  MoveL 2059 to (-200, -12.5, 57) mm, rotated rx 180 ry 0 rz 180 deg; joints [-15.333, -59.757, 128.123, 163.566, 69.173, -84.013]
  MoveL 2060 to (0, -12.5, 57) mm, rotated rx 180 ry 0 rz 180 deg; joints [-13.182, -51.64, 111.998, 164.918, 61.214, -82.606]
  MoveL 2061 to (0, -11.9, 57) mm, rotated rx 180 ry 0 rz 180 deg; joints [-13.182, -51.608, 111.999, 164.923, 61.246, -82.616]
  MoveL 2062 to (-200, -11.9, 57) mm, rotated rx 180 ry 0 rz 180 deg; joints [-15.333, -59.718, 128.125, 163.57, 69.212, -84.025]
  MoveL 2063 to (-200, -11.3, 57) mm, rotated rx 180 ry 0 rz 180 deg; joints [-15.333, -59.679, 128.126, 163.574, 69.251, -84.038]
  MoveL 2064 to (0, -11.3, 57) mm, rotated rx 180 ry 0 rz 180 deg; joints [-13.182, -51.576, 112.001, 164.927, 61.278, -82.626]
  MoveL 2065 to (0, -10.7, 57) mm, rotated rx 180 ry 0 rz 180 deg; joints [-13.182, -51.544, 112.002, 164.932, 61.31, -82.636]
  MoveL 2066 to (-200, -10.7, 57) mm, rotated rx 180 ry 0 rz 180 deg; joints [-15.333, -59.64, 128.127, 163.579, 69.289, -84.05]
  MoveL 2067 to (-200, -10.1, 57) mm, rotated rx 180 ry 0 rz 180 deg; joints [-15.333, -59.601, 128.129, 163.583, 69.328, -84.062]
  MoveL 2068 to (0, -10.1, 57) mm, rotated rx 180 ry 0 rz 180 deg; joints [-13.182, -51.512, 112.003, 164.937, 61.341, -82.645]
  MoveL 2069 to (0, -9.5, 57) mm, rotated rx 180 ry 0 rz 180 deg; joints [-13.182, -51.48, 112.004, 164.942, 61.373, -82.655]
  MoveL 2070 to (-200, -9.5, 57) mm, rotated rx 180 ry 0 rz 180 deg; joints [-15.333, -59.561, 128.13, 163.587, 69.367, -84.074]
  MoveL 2071 to (-200, -8.9, 57) mm, rotated rx 180 ry 0 rz 180 deg; joints [-15.333, -59.522, 128.131, 163.592, 69.406, -84.086]
  MoveL 2072 to (0, -8.9, 57) mm, rotated rx 180 ry 0 rz 180 deg; joints [-13.182, -51.449, 112.005, 164.946, 61.405, -82.665]
  MoveL 2073 to (0, -8.3, 57) mm, rotated rx 180 ry 0 rz 180 deg; joints [-13.182, -51.417, 112.006, 164.951, 61.437, -82.675]
  MoveL 2074 to (-200, -8.3, 57) mm, rotated rx 180 ry 0 rz 180 deg; joints [-15.333, -59.483, 128.132, 163.596, 69.444, -84.098]
  MoveL 2075 to (-200, -7.7, 57) mm, rotated rx 180 ry 0 rz 180 deg; joints [-15.333, -59.444, 128.133, 163.6, 69.483, -84.111]
  MoveL 2076 to (0, -7.7, 57) mm, rotated rx 180 ry 0 rz 180 deg; joints [-13.182, -51.385, 112.007, 164.956, 61.469, -82.684]
  MoveL 2077 to (0, -7.1, 57) mm, rotated rx 180 ry 0 rz 180 deg; joints [-13.182, -51.353, 112.008, 164.96, 61.501, -82.694]
  MoveL 2078 to (-200, -7.1, 57) mm, rotated rx 180 ry 0 rz 180 deg; joints [-15.333, -59.405, 128.135, 163.604, 69.522, -84.123]
  MoveL 2079 to (-200, -6.5, 57) mm, rotated rx 180 ry 0 rz 180 deg; joints [-15.333, -59.366, 128.136, 163.609, 69.56, -84.135]
  MoveL 2080 to (0, -6.5, 57) mm, rotated rx 180 ry 0 rz 180 deg; joints [-13.182, -51.321, 112.009, 164.965, 61.533, -82.704]
  MoveL 2081 to (0, -5.9, 57) mm, rotated rx 180 ry 0 rz 180 deg; joints [-13.182, -51.289, 112.01, 164.969, 61.564, -82.714]
  MoveL 2082 to (-200, -5.9, 57) mm, rotated rx 180 ry 0 rz 180 deg; joints [-15.333, -59.327, 128.137, 163.613, 69.599, -84.147]
  MoveL 2083 to (-200, -5.3, 57) mm, rotated rx 180 ry 0 rz 180 deg; joints [-15.333, -59.287, 128.138, 163.617, 69.637, -84.159]
  MoveL 2084 to (0, -5.3, 57) mm, rotated rx 180 ry 0 rz 180 deg; joints [-13.182, -51.257, 112.011, 164.974, 61.596, -82.723]
  MoveL 2085 to (0, -4.7, 57) mm, rotated rx 180 ry 0 rz 180 deg; joints [-13.182, -51.225, 112.012, 164.979, 61.628, -82.733]
  MoveL 2086 to (-200, -4.7, 57) mm, rotated rx 180 ry 0 rz 180 deg; joints [-15.333, -59.248, 128.139, 163.621, 69.676, -84.171]
  MoveL 2087 to (-200, -4.1, 57) mm, rotated rx 180 ry 0 rz 180 deg; joints [-15.333, -59.209, 128.14, 163.626, 69.715, -84.183]
  MoveL 2088 to (0, -4.1, 57) mm, rotated rx 180 ry 0 rz 180 deg; joints [-13.182, -51.193, 112.013, 164.983, 61.66, -82.743]
  MoveL 2089 to (0, -3.5, 57) mm, rotated rx 180 ry 0 rz 180 deg; joints [-13.182, -51.161, 112.014, 164.988, 61.692, -82.752]
  MoveL 2090 to (-200, -3.5, 57) mm, rotated rx 180 ry 0 rz 180 deg; joints [-15.333, -59.17, 128.141, 163.63, 69.753, -84.195]
  MoveL 2091 to (-200, -2.9, 57) mm, rotated rx 180 ry 0 rz 180 deg; joints [-15.333, -59.13, 128.142, 163.634, 69.792, -84.207]
  MoveL 2092 to (0, -2.9, 57) mm, rotated rx 180 ry 0 rz 180 deg; joints [-13.182, -51.129, 112.015, 164.992, 61.723, -82.762]
  MoveL 2093 to (0, -2.3, 57) mm, rotated rx 180 ry 0 rz 180 deg; joints [-13.182, -51.097, 112.015, 164.997, 61.755, -82.772]
  MoveL 2094 to (-200, -2.3, 57) mm, rotated rx 180 ry 0 rz 180 deg; joints [-15.333, -59.091, 128.142, 163.638, 69.83, -84.22]
  MoveL 2095 to (-200, -1.7, 57) mm, rotated rx 180 ry 0 rz 180 deg; joints [-15.333, -59.052, 128.143, 163.642, 69.869, -84.232]
  MoveL 2096 to (0, -1.7, 57) mm, rotated rx 180 ry 0 rz 180 deg; joints [-13.182, -51.064, 112.016, 165.002, 61.787, -82.781]
  MoveL 2097 to (0, -1.1, 57) mm, rotated rx 180 ry 0 rz 180 deg; joints [-13.182, -51.032, 112.017, 165.006, 61.818, -82.791]
  MoveL 2098 to (-200, -1.1, 57) mm, rotated rx 180 ry 0 rz 180 deg; joints [-15.333, -59.012, 128.144, 163.646, 69.907, -84.244]
  MoveL 2099 to (-200, -0.5, 57) mm, rotated rx 180 ry 0 rz 180 deg; joints [-15.333, -58.973, 128.145, 163.651, 69.946, -84.256]
  MoveL 2100 to (0, -0.5, 57) mm, rotated rx 180 ry 0 rz 180 deg; joints [-13.182, -51, 112.017, 165.011, 61.85, -82.801]
  MoveL 2101 to (0, 0, 57) mm, rotated rx 180 ry 0 rz 180 deg; joints [-13.182, -50.974, 112.018, 165.014, 61.876, -82.809]
  MoveL 2102 to (-200, 0, 57) mm, rotated rx 180 ry 0 rz 180 deg; joints [-15.333, -58.94, 128.145, 163.654, 69.978, -84.266]
  MoveL 2103 to (-200, 0, 57.4) mm, rotated rx 180 ry 0 rz 180 deg; joints [-15.351, -58.936, 128.137, 163.634, 69.976, -84.258]
  MoveL 2104 to (0, 0, 57.4) mm, rotated rx 180 ry 0 rz 180 deg; joints [-13.198, -50.97, 112.01, 164.996, 61.875, -82.799]
  MoveL 2105 to (0, -0.6, 57.4) mm, rotated rx 180 ry 0 rz 180 deg; joints [-13.198, -51.002, 112.009, 164.992, 61.843, -82.789]
  MoveL 2106 to (-200, -0.6, 57.4) mm, rotated rx 180 ry 0 rz 180 deg; joints [-15.351, -58.975, 128.136, 163.63, 69.937, -84.246]
  MoveL 2107 to (-200, -1.2, 57.4) mm, rotated rx 180 ry 0 rz 180 deg; joints [-15.351, -59.015, 128.135, 163.626, 69.899, -84.234]
  MoveL 2108 to (0, -1.2, 57.4) mm, rotated rx 180 ry 0 rz 180 deg; joints [-13.198, -51.034, 112.009, 164.987, 61.811, -82.78]
  MoveL 2109 to (0, -1.8, 57.4) mm, rotated rx 180 ry 0 rz 180 deg; joints [-13.198, -51.066, 112.008, 164.982, 61.78, -82.77]
  MoveL 2110 to (-200, -1.8, 57.4) mm, rotated rx 180 ry 0 rz 180 deg; joints [-15.351, -59.054, 128.135, 163.622, 69.86, -84.222]
  MoveL 2111 to (-200, -2.4, 57.4) mm, rotated rx 180 ry 0 rz 180 deg; joints [-15.351, -59.093, 128.134, 163.618, 69.822, -84.21]
  MoveL 2112 to (0, -2.4, 57.4) mm, rotated rx 180 ry 0 rz 180 deg; joints [-13.198, -51.098, 112.007, 164.978, 61.748, -82.76]
  MoveL 2113 to (0, -3, 57.4) mm, rotated rx 180 ry 0 rz 180 deg; joints [-13.198, -51.13, 112.006, 164.973, 61.716, -82.751]
  MoveL 2114 to (-200, -3, 57.4) mm, rotated rx 180 ry 0 rz 180 deg; joints [-15.351, -59.133, 128.133, 163.614, 69.783, -84.198]
  MoveL 2115 to (-200, -3.6, 57.4) mm, rotated rx 180 ry 0 rz 180 deg; joints [-15.351, -59.172, 128.132, 163.609, 69.744, -84.185]
  MoveL 2116 to (0, -3.6, 57.4) mm, rotated rx 180 ry 0 rz 180 deg; joints [-13.198, -51.162, 112.006, 164.969, 61.684, -82.741]
  MoveL 2117 to (0, -4.2, 57.4) mm, rotated rx 180 ry 0 rz 180 deg; joints [-13.198, -51.194, 112.005, 164.964, 61.653, -82.731]
  MoveL 2118 to (-200, -4.2, 57.4) mm, rotated rx 180 ry 0 rz 180 deg; joints [-15.351, -59.211, 128.131, 163.605, 69.706, -84.173]
  MoveL 2119 to (-200, -4.8, 57.4) mm, rotated rx 180 ry 0 rz 180 deg; joints [-15.351, -59.25, 128.13, 163.601, 69.667, -84.161]
  MoveL 2120 to (0, -4.8, 57.4) mm, rotated rx 180 ry 0 rz 180 deg; joints [-13.198, -51.226, 112.004, 164.96, 61.621, -82.722]
  MoveL 2121 to (0, -5.4, 57.4) mm, rotated rx 180 ry 0 rz 180 deg; joints [-13.198, -51.258, 112.003, 164.955, 61.589, -82.712]
  MoveL 2122 to (-200, -5.4, 57.4) mm, rotated rx 180 ry 0 rz 180 deg; joints [-15.351, -59.29, 128.129, 163.597, 69.629, -84.149]
  MoveL 2123 to (-200, -6, 57.4) mm, rotated rx 180 ry 0 rz 180 deg; joints [-15.351, -59.329, 128.128, 163.593, 69.59, -84.137]
  MoveL 2124 to (0, -6, 57.4) mm, rotated rx 180 ry 0 rz 180 deg; joints [-13.198, -51.29, 112.002, 164.95, 61.557, -82.702]
  MoveL 2125 to (0, -6.6, 57.4) mm, rotated rx 180 ry 0 rz 180 deg; joints [-13.198, -51.322, 112.001, 164.946, 61.525, -82.693]
  MoveL 2126 to (-200, -6.6, 57.4) mm, rotated rx 180 ry 0 rz 180 deg; joints [-15.351, -59.368, 128.127, 163.588, 69.551, -84.125]
  MoveL 2127 to (-200, -7.2, 57.4) mm, rotated rx 180 ry 0 rz 180 deg; joints [-15.351, -59.407, 128.126, 163.584, 69.513, -84.113]
  MoveL 2128 to (0, -7.2, 57.4) mm, rotated rx 180 ry 0 rz 180 deg; joints [-13.198, -51.354, 112, 164.941, 61.494, -82.683]
  MoveL 2129 to (0, -7.8, 57.4) mm, rotated rx 180 ry 0 rz 180 deg; joints [-13.198, -51.386, 111.999, 164.936, 61.462, -82.673]
  MoveL 2130 to (-200, -7.8, 57.4) mm, rotated rx 180 ry 0 rz 180 deg; joints [-15.351, -59.446, 128.125, 163.58, 69.474, -84.101]
  MoveL 2131 to (-200, -8.4, 57.4) mm, rotated rx 180 ry 0 rz 180 deg; joints [-15.351, -59.486, 128.124, 163.575, 69.436, -84.088]
  MoveL 2132 to (0, -8.4, 57.4) mm, rotated rx 180 ry 0 rz 180 deg; joints [-13.198, -51.418, 111.998, 164.932, 61.43, -82.663]
  MoveL 2133 to (0, -9, 57.4) mm, rotated rx 180 ry 0 rz 180 deg; joints [-13.198, -51.45, 111.997, 164.927, 61.398, -82.654]
  MoveL 2134 to (-200, -9, 57.4) mm, rotated rx 180 ry 0 rz 180 deg; joints [-15.351, -59.525, 128.123, 163.571, 69.397, -84.076]
  MoveL 2135 to (-200, -9.6, 57.4) mm, rotated rx 180 ry 0 rz 180 deg; joints [-15.351, -59.564, 128.121, 163.567, 69.358, -84.064]
  MoveL 2136 to (0, -9.6, 57.4) mm, rotated rx 180 ry 0 rz 180 deg; joints [-13.198, -51.482, 111.996, 164.922, 61.366, -82.644]
  MoveL 2137 to (0, -10.2, 57.4) mm, rotated rx 180 ry 0 rz 180 deg; joints [-13.198, -51.514, 111.995, 164.918, 61.334, -82.634]
  MoveL 2138 to (-200, -10.2, 57.4) mm, rotated rx 180 ry 0 rz 180 deg; joints [-15.351, -59.603, 128.12, 163.563, 69.319, -84.052]
  MoveL 2139 to (-200, -10.8, 57.4) mm, rotated rx 180 ry 0 rz 180 deg; joints [-15.351, -59.642, 128.119, 163.558, 69.281, -84.04]
  MoveL 2140 to (0, -10.8, 57.4) mm, rotated rx 180 ry 0 rz 180 deg; joints [-13.198, -51.546, 111.994, 164.913, 61.302, -82.624]
  MoveL 2141 to (0, -11.4, 57.4) mm, rotated rx 180 ry 0 rz 180 deg; joints [-13.198, -51.577, 111.992, 164.908, 61.27, -82.614]
  MoveL 2142 to (-200, -11.4, 57.4) mm, rotated rx 180 ry 0 rz 180 deg; joints [-15.351, -59.681, 128.117, 163.554, 69.242, -84.027]
  MoveL 2143 to (-200, -12, 57.4) mm, rotated rx 180 ry 0 rz 180 deg; joints [-15.351, -59.72, 128.116, 163.55, 69.203, -84.015]
  MoveL 2144 to (0, -12, 57.4) mm, rotated rx 180 ry 0 rz 180 deg; joints [-13.198, -51.609, 111.991, 164.903, 61.239, -82.605]
  MoveL 2145 to (0, -12.6, 57.4) mm, rotated rx 180 ry 0 rz 180 deg; joints [-13.198, -51.641, 111.99, 164.899, 61.207, -82.595]
  MoveL 2146 to (-200, -12.6, 57.4) mm, rotated rx 180 ry 0 rz 180 deg; joints [-15.351, -59.759, 128.115, 163.545, 69.164, -84.003]
  MoveL 2147 to (-200, -13.2, 57.4) mm, rotated rx 180 ry 0 rz 180 deg; joints [-15.351, -59.798, 128.113, 163.541, 69.126, -83.991]
  MoveL 2148 to (0, -13.2, 57.4) mm, rotated rx 180 ry 0 rz 180 deg; joints [-13.198, -51.673, 111.989, 164.894, 61.175, -82.585]
  MoveL 2149 to (0, -13.8, 57.4) mm, rotated rx 180 ry 0 rz 180 deg; joints [-13.198, -51.705, 111.987, 164.889, 61.143, -82.575]
  MoveL 2150 to (-200, -13.8, 57.4) mm, rotated rx 180 ry 0 rz 180 deg; joints [-15.351, -59.837, 128.112, 163.537, 69.087, -83.978]
  MoveL 2151 to (-200, -14.4, 57.4) mm, rotated rx 180 ry 0 rz 180 deg; joints [-15.351, -59.876, 128.11, 163.532, 69.048, -83.966]
  MoveL 2152 to (0, -14.4, 57.4) mm, rotated rx 180 ry 0 rz 180 deg; joints [-13.198, -51.736, 111.986, 164.884, 61.111, -82.565]
  MoveL 2153 to (0, -15, 57.4) mm, rotated rx 180 ry 0 rz 180 deg; joints [-13.198, -51.768, 111.985, 164.88, 61.079, -82.555]
  MoveL 2154 to (-200, -15, 57.4) mm, rotated rx 180 ry 0 rz 180 deg; joints [-15.351, -59.915, 128.109, 163.528, 69.009, -83.954]
  MoveL 2155 to (-200, -15.6, 57.4) mm, rotated rx 180 ry 0 rz 180 deg; joints [-15.351, -59.954, 128.107, 163.523, 68.97, -83.941]
  MoveL 2156 to (0, -15.6, 57.4) mm, rotated rx 180 ry 0 rz 180 deg; joints [-13.198, -51.8, 111.983, 164.875, 61.047, -82.545]
  MoveL 2157 to (0, -16.2, 57.4) mm, rotated rx 180 ry 0 rz 180 deg; joints [-13.198, -51.832, 111.982, 164.87, 61.015, -82.535]
  MoveL 2158 to (-200, -16.2, 57.4) mm, rotated rx 180 ry 0 rz 180 deg; joints [-15.351, -59.993, 128.106, 163.519, 68.932, -83.929]
  MoveL 2159 to (-200, -16.8, 57.4) mm, rotated rx 180 ry 0 rz 180 deg; joints [-15.351, -60.032, 128.104, 163.514, 68.893, -83.917]
  MoveL 2160 to (0, -16.8, 57.4) mm, rotated rx 180 ry 0 rz 180 deg; joints [-13.198, -51.863, 111.98, 164.865, 60.983, -82.526]
  MoveL 2161 to (0, -17.4, 57.4) mm, rotated rx 180 ry 0 rz 180 deg; joints [-13.198, -51.895, 111.979, 164.861, 60.951, -82.516]
  MoveL 2162 to (-200, -17.4, 57.4) mm, rotated rx 180 ry 0 rz 180 deg; joints [-15.351, -60.071, 128.102, 163.51, 68.854, -83.905]
  MoveL 2163 to (-200, -18, 57.4) mm, rotated rx 180 ry 0 rz 180 deg; joints [-15.351, -60.11, 128.101, 163.506, 68.815, -83.892]
  MoveL 2164 to (0, -18, 57.4) mm, rotated rx 180 ry 0 rz 180 deg; joints [-13.198, -51.927, 111.977, 164.856, 60.919, -82.506]
  MoveL 2165 to (0, -18.6, 57.4) mm, rotated rx 180 ry 0 rz 180 deg; joints [-13.198, -51.959, 111.976, 164.851, 60.886, -82.496]
  MoveL 2166 to (-200, -18.6, 57.4) mm, rotated rx 180 ry 0 rz 180 deg; joints [-15.351, -60.148, 128.099, 163.501, 68.776, -83.88]
  MoveL 2167 to (-200, -19.2, 57.4) mm, rotated rx 180 ry 0 rz 180 deg; joints [-15.351, -60.187, 128.097, 163.497, 68.737, -83.867]
  MoveL 2168 to (0, -19.2, 57.4) mm, rotated rx 180 ry 0 rz 180 deg; joints [-13.198, -51.99, 111.974, 164.846, 60.854, -82.486]
  MoveL 2169 to (0, -19.8, 57.4) mm, rotated rx 180 ry 0 rz 180 deg; joints [-13.198, -52.022, 111.972, 164.841, 60.822, -82.476]
  MoveL 2170 to (-200, -19.8, 57.4) mm, rotated rx 180 ry 0 rz 180 deg; joints [-15.351, -60.226, 128.095, 163.492, 68.698, -83.855]
  MoveL 2171 to (-200, -20.4, 57.4) mm, rotated rx 180 ry 0 rz 180 deg; joints [-15.351, -60.265, 128.094, 163.488, 68.659, -83.843]
  MoveL 2172 to (0, -20.4, 57.4) mm, rotated rx 180 ry 0 rz 180 deg; joints [-13.198, -52.053, 111.971, 164.836, 60.79, -82.466]
  MoveL 2173 to (0, -21, 57.4) mm, rotated rx 180 ry 0 rz 180 deg; joints [-13.198, -52.085, 111.969, 164.831, 60.758, -82.456]
  MoveL 2174 to (-200, -21, 57.4) mm, rotated rx 180 ry 0 rz 180 deg; joints [-15.351, -60.304, 128.092, 163.483, 68.62, -83.83]
  MoveL 2175 to (-200, -21.6, 57.4) mm, rotated rx 180 ry 0 rz 180 deg; joints [-15.351, -60.342, 128.09, 163.479, 68.581, -83.818]
  MoveL 2176 to (0, -21.6, 57.4) mm, rotated rx 180 ry 0 rz 180 deg; joints [-13.198, -52.117, 111.967, 164.827, 60.726, -82.446]
  MoveL 2177 to (0, -22.2, 57.4) mm, rotated rx 180 ry 0 rz 180 deg; joints [-13.198, -52.148, 111.966, 164.822, 60.694, -82.436]
  MoveL 2178 to (-200, -22.2, 57.4) mm, rotated rx 180 ry 0 rz 180 deg; joints [-15.351, -60.381, 128.088, 163.474, 68.542, -83.805]
  MoveL 2179 to (-200, -22.8, 57.4) mm, rotated rx 180 ry 0 rz 180 deg; joints [-15.351, -60.42, 128.086, 163.469, 68.503, -83.793]
  MoveL 2180 to (0, -22.8, 57.4) mm, rotated rx 180 ry 0 rz 180 deg; joints [-13.198, -52.18, 111.964, 164.817, 60.662, -82.426]
  MoveL 2181 to (0, -23.4, 57.4) mm, rotated rx 180 ry 0 rz 180 deg; joints [-13.198, -52.211, 111.962, 164.812, 60.629, -82.416]
  MoveL 2182 to (-200, -23.4, 57.4) mm, rotated rx 180 ry 0 rz 180 deg; joints [-15.351, -60.459, 128.084, 163.465, 68.464, -83.781]
  MoveL 2183 to (-200, -24, 57.4) mm, rotated rx 180 ry 0 rz 180 deg; joints [-15.351, -60.497, 128.082, 163.46, 68.425, -83.768]
  MoveL 2184 to (0, -24, 57.4) mm, rotated rx 180 ry 0 rz 180 deg; joints [-13.198, -52.243, 111.96, 164.807, 60.597, -82.406]
  MoveL 2185 to (0, -24.6, 57.4) mm, rotated rx 180 ry 0 rz 180 deg; joints [-13.198, -52.274, 111.958, 164.802, 60.565, -82.396]
  MoveL 2186 to (-200, -24.6, 57.4) mm, rotated rx 180 ry 0 rz 180 deg; joints [-15.351, -60.536, 128.08, 163.456, 68.386, -83.756]
  MoveL 2187 to (-200, -25.2, 57.4) mm, rotated rx 180 ry 0 rz 180 deg; joints [-15.351, -60.575, 128.078, 163.451, 68.347, -83.743]
  MoveL 2188 to (0, -25.2, 57.4) mm, rotated rx 180 ry 0 rz 180 deg; joints [-13.198, -52.306, 111.957, 164.797, 60.533, -82.386]
  MoveL 2189 to (0, -25.8, 57.4) mm, rotated rx 180 ry 0 rz 180 deg; joints [-13.198, -52.337, 111.955, 164.792, 60.501, -82.376]
  MoveL 2190 to (-200, -25.8, 57.4) mm, rotated rx 180 ry 0 rz 180 deg; joints [-15.351, -60.613, 128.076, 163.447, 68.308, -83.731]
  MoveL 2191 to (-200, -26.4, 57.4) mm, rotated rx 180 ry 0 rz 180 deg; joints [-15.351, -60.652, 128.073, 163.442, 68.269, -83.718]
  MoveL 2192 to (0, -26.4, 57.4) mm, rotated rx 180 ry 0 rz 180 deg; joints [-13.198, -52.369, 111.953, 164.787, 60.468, -82.366]
  MoveL 2193 to (0, -27, 57.4) mm, rotated rx 180 ry 0 rz 180 deg; joints [-13.198, -52.4, 111.951, 164.782, 60.436, -82.356]
  MoveL 2194 to (-200, -27, 57.4) mm, rotated rx 180 ry 0 rz 180 deg; joints [-15.351, -60.69, 128.071, 163.437, 68.23, -83.706]
  MoveL 2195 to (-200, -27.6, 57.4) mm, rotated rx 180 ry 0 rz 180 deg; joints [-15.351, -60.729, 128.069, 163.433, 68.191, -83.693]
  MoveL 2196 to (0, -27.6, 57.4) mm, rotated rx 180 ry 0 rz 180 deg; joints [-13.198, -52.432, 111.949, 164.777, 60.404, -82.346]
  MoveL 2197 to (0, -28.2, 57.4) mm, rotated rx 180 ry 0 rz 180 deg; joints [-13.198, -52.463, 111.947, 164.772, 60.372, -82.335]
  MoveL 2198 to (-200, -28.2, 57.4) mm, rotated rx 180 ry 0 rz 180 deg; joints [-15.351, -60.768, 128.067, 163.428, 68.152, -83.681]
  MoveL 2199 to (-200, -28.8, 57.4) mm, rotated rx 180 ry 0 rz 180 deg; joints [-15.351, -60.806, 128.065, 163.423, 68.113, -83.668]
  MoveL 2200 to (0, -28.8, 57.4) mm, rotated rx 180 ry 0 rz 180 deg; joints [-13.198, -52.495, 111.945, 164.767, 60.339, -82.325]
  MoveL 2201 to (0, -29.4, 57.4) mm, rotated rx 180 ry 0 rz 180 deg; joints [-13.198, -52.526, 111.943, 164.762, 60.307, -82.315]
  MoveL 2202 to (-200, -29.4, 57.4) mm, rotated rx 180 ry 0 rz 180 deg; joints [-15.351, -60.845, 128.062, 163.419, 68.074, -83.655]
  MoveL 2203 to (-200, -30, 57.4) mm, rotated rx 180 ry 0 rz 180 deg; joints [-15.351, -60.883, 128.06, 163.414, 68.034, -83.643]
  MoveL 2204 to (0, -30, 57.4) mm, rotated rx 180 ry 0 rz 180 deg; joints [-13.198, -52.557, 111.94, 164.757, 60.275, -82.305]
  MoveL 2205 to (0, -30.6, 57.38) mm, rotated rx 177.23 ry 0 rz 180 deg; joints [-13.263, -53.471, 111.83, 164.524, 59.296, -84.725]
  MoveL 2206 to (-200, -30.6, 57.38) mm, rotated rx 177.23 ry 0 rz 180 deg; joints [-15.426, -62.007, 127.939, 163.184, 66.851, -85.997]
  MoveL 2207 to (-200, -31.2, 57.34) mm, rotated rx 174.45 ry 0 rz 180 deg; joints [-15.462, -63.127, 127.807, 162.985, 65.658, -88.356]
  MoveL 2208 to (0, -31.2, 57.34) mm, rotated rx 174.45 ry 0 rz 180 deg; joints [-13.295, -54.381, 111.71, 164.32, 58.308, -87.156]
  MoveL 2209 to (0, -31.79, 57.27) mm, rotated rx 171.68 ry 0 rz 180 deg; joints [-13.291, -55.286, 111.581, 164.147, 57.312, -89.598]
  MoveL 2210 to (-200, -31.79, 57.27) mm, rotated rx 171.68 ry 0 rz 180 deg; joints [-15.458, -64.238, 127.664, 162.818, 64.458, -90.723]
  MoveL 2211 to (-200, -32.38, 57.17) mm, rotated rx 168.91 ry 0 rz 180 deg; joints [-15.415, -65.34, 127.51, 162.683, 63.253, -93.102]
  MoveL 2212 to (0, -32.38, 57.17) mm, rotated rx 168.91 ry 0 rz 180 deg; joints [-13.253, -56.184, 111.442, 164.006, 56.31, -92.056]
  MoveL 2213 to (0, -32.97, 57.04) mm, rotated rx 166.14 ry 0 rz 180 deg; joints [-13.181, -57.072, 111.295, 163.898, 55.304, -94.531]
  MoveL 2214 to (-200, -32.97, 57.04) mm, rotated rx 166.14 ry 0 rz 180 deg; joints [-15.332, -66.429, 127.346, 162.582, 62.045, -95.496]
  MoveL 2215 to (-200, -33.55, 56.88) mm, rotated rx 163.37 ry 0 rz 180 deg; joints [-15.209, -67.502, 127.171, 162.516, 60.837, -97.908]
  MoveL 2216 to (0, -33.55, 56.88) mm, rotated rx 163.37 ry 0 rz 180 deg; joints [-13.074, -57.948, 111.14, 163.825, 54.296, -97.026]
  MoveL 2217 to (0, -34.12, 56.7) mm, rotated rx 160.59 ry 0 rz 180 deg; joints [-12.934, -58.811, 110.977, 163.787, 53.287, -99.546]
  MoveL 2218 to (-200, -34.12, 56.7) mm, rotated rx 160.59 ry 0 rz 180 deg; joints [-15.048, -68.558, 126.988, 162.487, 59.629, -100.343]
  MoveL 2219 to (-200, -34.68, 56.48) mm, rotated rx 157.82 ry 0 rz 180 deg; joints [-14.847, -69.594, 126.795, 162.497, 58.426, -102.803]
  MoveL 2220 to (0, -34.68, 56.48) mm, rotated rx 157.82 ry 0 rz 180 deg; joints [-12.759, -59.658, 110.807, 163.788, 52.28, -102.092]
  MoveL 2221 to (0, -35.23, 56.24) mm, rotated rx 155.05 ry 0 rz 180 deg; joints [-12.551, -60.488, 110.631, 163.828, 51.277, -104.668]
  MoveL 2222 to (-200, -35.23, 56.24) mm, rotated rx 155.05 ry 0 rz 180 deg; joints [-14.607, -70.608, 126.596, 162.547, 57.229, -105.293]
  MoveL 2223 to (-200, -35.77, 55.98) mm, rotated rx 152.28 ry 0 rz 180 deg; joints [-14.329, -71.597, 126.389, 162.64, 56.039, -107.818]
  MoveL 2224 to (0, -35.77, 55.98) mm, rotated rx 152.28 ry 0 rz 180 deg; joints [-12.309, -61.299, 110.448, 163.909, 50.279, -107.279]
  MoveL 2225 to (0, -36.29, 55.69) mm, rotated rx 149.5 ry 0 rz 180 deg; joints [-12.034, -62.089, 110.261, 164.035, 49.289, -109.926]
  MoveL 2226 to (-200, -36.29, 55.69) mm, rotated rx 149.5 ry 0 rz 180 deg; joints [-14.012, -72.561, 126.176, 162.777, 54.861, -110.38]
  MoveL 2227 to (-200, -36.8, 55.37) mm, rotated rx 146.73 ry 0 rz 180 deg; joints [-13.658, -73.496, 125.958, 162.962, 53.696, -112.985]
  MoveL 2228 to (0, -36.8, 55.37) mm, rotated rx 146.73 ry 0 rz 180 deg; joints [-11.727, -62.857, 110.069, 164.206, 48.309, -112.614]
  MoveL 2229 to (0, -37.3, 55.03) mm, rotated rx 143.96 ry 0 rz 180 deg; joints [-11.388, -63.601, 109.874, 164.426, 47.342, -115.346]
  MoveL 2230 to (-200, -37.3, 55.03) mm, rotated rx 143.96 ry 0 rz 180 deg; joints [-13.267, -74.401, 125.735, 163.197, 52.547, -115.635]
  MoveL 2231 to (-200, -37.77, 54.66) mm, rotated rx 141.19 ry 0 rz 180 deg; joints [-12.839, -75.275, 125.51, 163.485, 51.417, -118.337]
  MoveL 2232 to (0, -37.77, 54.66) mm, rotated rx 141.19 ry 0 rz 180 deg; joints [-11.017, -64.32, 109.676, 164.696, 46.39, -118.125]
  MoveL 2233 to (0, -38.23, 54.27) mm, rotated rx 138.41 ry 0 rz 180 deg; joints [-10.616, -65.012, 109.477, 165.02, 45.455, -120.955]
  MoveL 2234 to (-200, -38.23, 54.27) mm, rotated rx 138.41 ry 0 rz 180 deg; joints [-12.376, -76.116, 125.283, 163.828, 50.308, -121.093]
  MoveL 2235 to (-200, -38.67, 53.87) mm, rotated rx 135.64 ry 0 rz 180 deg; joints [-11.877, -76.921, 125.054, 164.23, 49.223, -123.908]
  MoveL 2236 to (0, -38.67, 53.87) mm, rotated rx 135.64 ry 0 rz 180 deg; joints [-10.185, -65.676, 109.276, 165.398, 44.54, -123.839]
  MoveL 2237 to (0, -39.09, 53.44) mm, rotated rx 132.87 ry 0 rz 180 deg; joints [-9.724, -66.311, 109.076, 165.835, 43.648, -126.78]
  MoveL 2238 to (-200, -39.09, 53.44) mm, rotated rx 132.87 ry 0 rz 180 deg; joints [-11.344, -77.69, 124.826, 164.693, 48.166, -126.785]
  MoveL 2239 to (-200, -39.48, 52.99) mm, rotated rx 130.1 ry 0 rz 180 deg; joints [-10.777, -78.422, 124.599, 165.221, 47.14, -129.729]
  MoveL 2240 to (0, -39.48, 52.99) mm, rotated rx 130.1 ry 0 rz 180 deg; joints [-9.235, -66.915, 108.876, 166.332, 42.781, -129.783]
  MoveL 2241 to (0, -39.86, 52.52) mm, rotated rx 127.33 ry 0 rz 180 deg; joints [-8.72, -67.488, 108.679, 166.89, 41.942, -132.848]
  MoveL 2242 to (-200, -39.86, 52.52) mm, rotated rx 127.33 ry 0 rz 180 deg; joints [-10.179, -79.115, 124.375, 165.815, 46.147, -132.742]
  MoveL 2243 to (-200, -40.21, 52.03) mm, rotated rx 124.55 ry 0 rz 180 deg; joints [-9.549, -79.768, 124.154, 166.478, 45.192, -135.829]
  MoveL 2244 to (0, -40.21, 52.03) mm, rotated rx 124.55 ry 0 rz 180 deg; joints [-8.177, -68.028, 108.485, 167.513, 41.135, -135.979]
  MoveL 2245 to (0, -40.54, 51.53) mm, rotated rx 121.78 ry 0 rz 180 deg; joints [-7.61, -68.534, 108.294, 168.2, 40.362, -139.176]
  MoveL 2246 to (-200, -40.54, 51.53) mm, rotated rx 121.78 ry 0 rz 180 deg; joints [-8.89, -80.379, 123.938, 167.212, 44.278, -138.99]
  MoveL 2247 to (-200, -40.84, 51.01) mm, rotated rx 119.01 ry 0 rz 180 deg; joints [-8.202, -80.948, 123.727, 168.018, 43.409, -142.228]
  MoveL 2248 to (0, -40.84, 51.01) mm, rotated rx 119.01 ry 0 rz 180 deg; joints [-7.019, -69.006, 108.108, 168.954, 39.627, -142.441]
  MoveL 2249 to (0, -41.12, 50.48) mm, rotated rx 116.23 ry 0 rz 180 deg; joints [-6.405, -69.443, 107.928, 169.774, 38.933, -145.777]
  MoveL 2250 to (-200, -41.12, 50.48) mm, rotated rx 116.23 ry 0 rz 180 deg; joints [-7.487, -81.475, 123.523, 168.898, 42.587, -145.544]
  MoveL 2251 to (-200, -41.38, 49.94) mm, rotated rx 113.46 ry 0 rz 180 deg; joints [-6.747, -81.957, 123.327, 169.851, 41.819, -148.938]
  MoveL 2252 to (0, -41.38, 49.94) mm, rotated rx 113.46 ry 0 rz 180 deg; joints [-5.771, -69.843, 107.754, 170.66, 38.283, -149.18]
  MoveL 2253 to (0, -41.6, 49.38) mm, rotated rx 110.69 ry 0 rz 180 deg; joints [-5.117, -70.207, 107.588, 171.61, 37.679, -152.651]
  MoveL 2254 to (-200, -41.6, 49.38) mm, rotated rx 110.69 ry 0 rz 180 deg; joints [-5.984, -82.395, 123.14, 170.876, 41.107, -152.409]
  MoveL 2255 to (-200, -41.8, 48.81) mm, rotated rx 107.92 ry 0 rz 180 deg; joints [-5.199, -82.787, 122.963, 171.971, 40.454, -155.956]
  MoveL 2256 to (0, -41.8, 48.81) mm, rotated rx 107.92 ry 0 rz 180 deg; joints [-4.445, -70.533, 107.43, 172.623, 37.126, -156.188]
  MoveL 2257 to (0, -41.97, 48.24) mm, rotated rx 105.15 ry 0 rz 180 deg; joints [-3.756, -70.821, 107.281, 173.695, 36.626, -159.787]
  MoveL 2258 to (-200, -41.97, 48.24) mm, rotated rx 105.15 ry 0 rz 180 deg; joints [-4.395, -83.134, 122.796, 173.134, 39.865, -159.573]
  MoveL 2259 to (-200, -42.11, 47.66) mm, rotated rx 102.37 ry 0 rz 180 deg; joints [-3.573, -83.434, 122.641, 174.359, 39.343, -163.258]
  MoveL 2260 to (0, -42.11, 47.66) mm, rotated rx 102.37 ry 0 rz 180 deg; joints [-3.053, -71.071, 107.141, 174.824, 36.181, -163.445]
  MoveL 2261 to (0, -42.23, 47.07) mm, rotated rx 99.6 ry 0 rz 180 deg; joints [-2.337, -71.283, 107.012, 176.001, 35.796, -167.154]
  MoveL 2262 to (-200, -42.23, 47.07) mm, rotated rx 99.6 ry 0 rz 180 deg; joints [-2.736, -83.688, 122.498, 175.64, 38.891, -167.003]
  MoveL 2263 to (-200, -42.31, 46.47) mm, rotated rx 96.83 ry 0 rz 180 deg; joints [-1.886, -83.894, 122.368, 176.971, 38.512, -170.8]
  MoveL 2264 to (0, -42.31, 46.47) mm, rotated rx 96.83 ry 0 rz 180 deg; joints [-1.611, -71.455, 106.894, 177.223, 35.471, -170.909]
  MoveL 2265 to (0, -42.37, 45.88) mm, rotated rx 94.06 ry 0 rz 180 deg; joints [-0.875, -71.588, 106.787, 178.482, 35.208, -174.704]
  MoveL 2266 to (-200, -42.37, 45.88) mm, rotated rx 94.06 ry 0 rz 180 deg; joints [-1.024, -84.054, 122.251, 178.344, 38.209, -174.643]
  MoveL 2267 to (-200, -42.4, 45.28) mm, rotated rx 91.28 ry 0 rz 180 deg; joints [-0.155, -84.166, 122.148, 179.748, 37.983, -178.518]
  MoveL 2268 to (0, -42.4, 45.28) mm, rotated rx 91.28 ry 0 rz 180 deg; joints [-0.132, -71.682, 106.692, 179.769, 35.01, -178.527]
  MoveL 2269 to (0, -42.4, 44.68) mm, rotated rx 90 ry 0 rz 180 deg; joints [0.227, -71.712, 106.652, -179.604, 34.941, 179.675]
  MoveL 2270 to (-200, -42.4, 44.68) mm, rotated rx 90 ry 0 rz 180 deg; joints [0.266, -84.201, 122.105, -179.567, 37.905, 179.659]
  MoveL 2271 to (-200, -42.4, 44.08) mm, rotated rx 90 ry 0 rz 180 deg; joints [0.295, -84.201, 122.105, -179.52, 37.905, 179.621]
  MoveL 2272 to (0, -42.4, 44.08) mm, rotated rx 90 ry 0 rz 180 deg; joints [0.252, -71.711, 106.651, -179.56, 34.941, 179.639]
  MoveL 2273 to (0, -42.4, 43.48) mm, rotated rx 90 ry 0 rz 180 deg; joints [0.277, -71.711, 106.651, -179.516, 34.941, 179.603]
  MoveL 2274 to (-200, -42.4, 43.48) mm, rotated rx 90 ry 0 rz 180 deg; joints [0.324, -84.201, 122.105, -179.472, 37.905, 179.583]
  MoveL 2275 to (-200, -42.4, 42.88) mm, rotated rx 90 ry 0 rz 180 deg; joints [0.354, -84.201, 122.105, -179.424, 37.906, 179.546]
  MoveL 2276 to (0, -42.4, 42.88) mm, rotated rx 90 ry 0 rz 180 deg; joints [0.302, -71.711, 106.651, -179.472, 34.941, 179.568]
  MoveL 2277 to (0, -42.4, 42.28) mm, rotated rx 90 ry 0 rz 180 deg; joints [0.327, -71.711, 106.651, -179.429, 34.941, 179.532]
  MoveL 2278 to (-200, -42.4, 42.28) mm, rotated rx 90 ry 0 rz 180 deg; joints [0.383, -84.2, 122.104, -179.377, 37.906, 179.508]
  MoveL 2279 to (-200, -42.4, 41.68) mm, rotated rx 90 ry 0 rz 180 deg; joints [0.412, -84.2, 122.104, -179.329, 37.906, 179.47]
  MoveL 2280 to (0, -42.4, 41.68) mm, rotated rx 90 ry 0 rz 180 deg; joints [0.352, -71.711, 106.65, -179.385, 34.941, 179.496]
  MoveL 2281 to (0, -42.4, 41.08) mm, rotated rx 90 ry 0 rz 180 deg; joints [0.377, -71.71, 106.65, -179.341, 34.941, 179.46]
  MoveL 2282 to (-200, -42.4, 41.08) mm, rotated rx 90 ry 0 rz 180 deg; joints [0.442, -84.2, 122.104, -179.281, 37.906, 179.433]
  MoveL 2283 to (-200, -42.4, 40.48) mm, rotated rx 90 ry 0 rz 180 deg; joints [0.471, -84.199, 122.103, -179.233, 37.907, 179.395]
  MoveL 2284 to (0, -42.4, 40.48) mm, rotated rx 90 ry 0 rz 180 deg; joints [0.402, -71.71, 106.65, -179.297, 34.942, 179.424]
  MoveL 2285 to (0, -42.4, 39.88) mm, rotated rx 90 ry 0 rz 180 deg; joints [0.427, -71.71, 106.649, -179.254, 34.942, 179.388]
  MoveL 2286 to (-200, -42.4, 39.88) mm, rotated rx 90 ry 0 rz 180 deg; joints [0.5, -84.199, 122.103, -179.186, 37.907, 179.357]
  MoveL 2287 to (-200, -42.4, 39.28) mm, rotated rx 90 ry 0 rz 180 deg; joints [0.53, -84.199, 122.103, -179.138, 37.907, 179.32]
  MoveL 2288 to (0, -42.4, 39.28) mm, rotated rx 90 ry 0 rz 180 deg; joints [0.452, -71.71, 106.649, -179.21, 34.942, 179.352]
  MoveL 2289 to (0, -42.4, 38.68) mm, rotated rx 90 ry 0 rz 180 deg; joints [0.478, -71.709, 106.649, -179.166, 34.942, 179.317]
  MoveL 2290 to (-200, -42.4, 38.68) mm, rotated rx 90 ry 0 rz 180 deg; joints [0.559, -84.198, 122.102, -179.09, 37.907, 179.282]
  MoveL 2291 to (-200, -42.4, 38.08) mm, rotated rx 90 ry 0 rz 180 deg; joints [0.588, -84.198, 122.102, -179.042, 37.908, 179.244]
  MoveL 2292 to (0, -42.4, 38.08) mm, rotated rx 90 ry 0 rz 180 deg; joints [0.503, -71.709, 106.648, -179.122, 34.942, 179.281]
  MoveL 2293 to (0, -42.4, 37.48) mm, rotated rx 90 ry 0 rz 180 deg; joints [0.528, -71.709, 106.648, -179.079, 34.943, 179.245]
  MoveL 2294 to (-200, -42.4, 37.48) mm, rotated rx 90 ry 0 rz 180 deg; joints [0.618, -84.198, 122.101, -178.995, 37.908, 179.207]
  MoveL 2295 to (-200, -42.4, 36.88) mm, rotated rx 90 ry 0 rz 180 deg; joints [0.647, -84.197, 122.101, -178.947, 37.908, 179.169]
  MoveL 2296 to (0, -42.4, 36.88) mm, rotated rx 90 ry 0 rz 180 deg; joints [0.553, -71.708, 106.647, -179.035, 34.943, 179.209]
  MoveL 2297 to (0, -42.4, 36.28) mm, rotated rx 90 ry 0 rz 180 deg; joints [0.578, -71.708, 106.647, -178.991, 34.943, 179.173]
  MoveL 2298 to (-200, -42.4, 36.28) mm, rotated rx 90 ry 0 rz 180 deg; joints [0.676, -84.197, 122.1, -178.899, 37.909, 179.131]
  MoveL 2299 to (-200, -42.4, 35.68) mm, rotated rx 90 ry 0 rz 180 deg; joints [0.706, -84.196, 122.1, -178.851, 37.909, 179.094]
  MoveL 2300 to (0, -42.4, 35.68) mm, rotated rx 90 ry 0 rz 180 deg; joints [0.603, -71.708, 106.646, -178.948, 34.943, 179.137]
  MoveL 2301 to (0, -42.4, 35.08) mm, rotated rx 90 ry 0 rz 180 deg; joints [0.628, -71.707, 106.646, -178.904, 34.943, 179.101]
  MoveL 2302 to (-200, -42.4, 35.08) mm, rotated rx 90 ry 0 rz 180 deg; joints [0.735, -84.196, 122.099, -178.804, 37.91, 179.056]
  MoveL 2303 to (-200, -42.4, 34.48) mm, rotated rx 90 ry 0 rz 180 deg; joints [0.764, -84.195, 122.099, -178.756, 37.91, 179.018]
  MoveL 2304 to (0, -42.4, 34.48) mm, rotated rx 90 ry 0 rz 180 deg; joints [0.653, -71.707, 106.645, -178.86, 34.944, 179.065]
  MoveL 2305 to (0, -42.4, 33.88) mm, rotated rx 90 ry 0 rz 180 deg; joints [0.678, -71.706, 106.645, -178.816, 34.944, 179.03]
  MoveL 2306 to (-200, -42.4, 33.88) mm, rotated rx 90 ry 0 rz 180 deg; joints [0.794, -84.195, 122.098, -178.708, 37.911, 178.981]
  MoveL 2307 to (-200, -42.4, 33.28) mm, rotated rx 90 ry 0 rz 180 deg; joints [0.823, -84.194, 122.098, -178.661, 37.911, 178.943]
  MoveL 2308 to (0, -42.4, 33.28) mm, rotated rx 90 ry 0 rz 180 deg; joints [0.703, -71.706, 106.644, -178.773, 34.944, 178.994]
  MoveL 2309 to (0, -42.4, 32.68) mm, rotated rx 90 ry 0 rz 180 deg; joints [0.728, -71.705, 106.643, -178.729, 34.945, 178.958]
  MoveL 2310 to (-200, -42.4, 32.68) mm, rotated rx 90 ry 0 rz 180 deg; joints [0.852, -84.194, 122.097, -178.613, 37.912, 178.905]
  MoveL 2311 to (-200, -42.4, 32.08) mm, rotated rx 90 ry 0 rz 180 deg; joints [0.882, -84.193, 122.096, -178.565, 37.912, 178.868]
  MoveL 2312 to (0, -42.4, 32.08) mm, rotated rx 90 ry 0 rz 180 deg; joints [0.753, -71.705, 106.643, -178.685, 34.945, 178.922]
  MoveL 2313 to (0, -42.4, 31.48) mm, rotated rx 90 ry 0 rz 180 deg; joints [0.778, -71.704, 106.642, -178.641, 34.945, 178.886]
  MoveL 2314 to (-200, -42.4, 31.48) mm, rotated rx 90 ry 0 rz 180 deg; joints [0.911, -84.192, 122.096, -178.517, 37.913, 178.83]
  MoveL 2315 to (-200, -42.4, 30.88) mm, rotated rx 90 ry 0 rz 180 deg; joints [0.94, -84.192, 122.095, -178.47, 37.913, 178.793]
  MoveL 2316 to (0, -42.4, 30.88) mm, rotated rx 90 ry 0 rz 180 deg; joints [0.803, -71.704, 106.641, -178.598, 34.945, 178.85]
  MoveL 2317 to (0, -42.4, 30.28) mm, rotated rx 90 ry 0 rz 180 deg; joints [0.828, -71.703, 106.641, -178.554, 34.946, 178.815]
  MoveL 2318 to (-200, -42.4, 30.28) mm, rotated rx 90 ry 0 rz 180 deg; joints [0.97, -84.191, 122.094, -178.422, 37.914, 178.755]
  MoveL 2319 to (-200, -42.4, 29.68) mm, rotated rx 90 ry 0 rz 180 deg; joints [0.999, -84.19, 122.093, -178.374, 37.914, 178.717]
  MoveL 2320 to (0, -42.4, 29.68) mm, rotated rx 90 ry 0 rz 180 deg; joints [0.853, -71.703, 106.64, -178.51, 34.946, 178.779]
  MoveL 2321 to (0, -42.4, 29.08) mm, rotated rx 90 ry 0 rz 180 deg; joints [0.878, -71.702, 106.639, -178.466, 34.946, 178.743]
  MoveL 2322 to (-200, -42.4, 29.08) mm, rotated rx 90 ry 0 rz 180 deg; joints [1.028, -84.19, 122.093, -178.326, 37.915, 178.68]
  MoveL 2323 to (-200, -42.4, 28.48) mm, rotated rx 90 ry 0 rz 180 deg; joints [1.058, -84.189, 122.092, -178.279, 37.915, 178.642]
  MoveL 2324 to (0, -42.4, 28.48) mm, rotated rx 90 ry 0 rz 180 deg; joints [0.903, -71.702, 106.638, -178.423, 34.947, 178.707]
  MoveL 2325 to (0, -42.4, 27.88) mm, rotated rx 90 ry 0 rz 180 deg; joints [0.928, -71.701, 106.638, -178.379, 34.947, 178.671]
  MoveL 2326 to (-200, -42.4, 27.88) mm, rotated rx 90 ry 0 rz 180 deg; joints [1.087, -84.188, 122.091, -178.231, 37.916, 178.604]
  MoveL 2327 to (-200, -42.4, 27.28) mm, rotated rx 90 ry 0 rz 180 deg; joints [1.116, -84.188, 122.09, -178.183, 37.917, 178.567]
  MoveL 2328 to (0, -42.4, 27.28) mm, rotated rx 90 ry 0 rz 180 deg; joints [0.954, -71.701, 106.637, -178.335, 34.948, 178.635]
  MoveL 2329 to (0, -42.4, 26.68) mm, rotated rx 90 ry 0 rz 180 deg; joints [0.979, -71.7, 106.636, -178.291, 34.948, 178.599]
  MoveL 2330 to (-200, -42.4, 26.68) mm, rotated rx 90 ry 0 rz 180 deg; joints [1.146, -84.187, 122.089, -178.136, 37.917, 178.529]
  MoveL 2331 to (-200, -42.4, 26.08) mm, rotated rx 90 ry 0 rz 180 deg; joints [1.175, -84.186, 122.089, -178.088, 37.918, 178.491]
  MoveL 2332 to (0, -42.4, 26.08) mm, rotated rx 90 ry 0 rz 180 deg; joints [1.004, -71.699, 106.635, -178.248, 34.948, 178.564]
  MoveL 2333 to (0, -42.4, 25.48) mm, rotated rx 90 ry 0 rz 180 deg; joints [1.029, -71.699, 106.634, -178.204, 34.949, 178.528]
  MoveL 2334 to (-200, -42.4, 25.48) mm, rotated rx 90 ry 0 rz 180 deg; joints [1.204, -84.185, 122.088, -178.04, 37.919, 178.454]
  MoveL 2335 to (-200, -42.4, 24.88) mm, rotated rx 90 ry 0 rz 180 deg; joints [1.234, -84.184, 122.087, -177.993, 37.919, 178.416]
  MoveL 2336 to (0, -42.4, 24.88) mm, rotated rx 90 ry 0 rz 180 deg; joints [1.054, -71.698, 106.633, -178.16, 34.949, 178.492]
  MoveL 2337 to (0, -42.4, 24.28) mm, rotated rx 90 ry 0 rz 180 deg; joints [1.079, -71.697, 106.632, -178.117, 34.95, 178.456]
  MoveL 2338 to (-200, -42.4, 24.28) mm, rotated rx 90 ry 0 rz 180 deg; joints [1.263, -84.184, 122.086, -177.945, 37.92, 178.379]
  MoveL 2339 to (-200, -42.4, 23.68) mm, rotated rx 90 ry 0 rz 180 deg; joints [1.292, -84.183, 122.085, -177.897, 37.921, 178.341]
  MoveL 2340 to (0, -42.4, 23.68) mm, rotated rx 90 ry 0 rz 180 deg; joints [1.104, -71.697, 106.631, -178.073, 34.95, 178.42]
  MoveL 2341 to (0, -42.4, 23.08) mm, rotated rx 90 ry 0 rz 180 deg; joints [1.129, -71.696, 106.63, -178.029, 34.95, 178.384]
  MoveL 2342 to (-200, -42.4, 23.08) mm, rotated rx 90 ry 0 rz 180 deg; joints [1.321, -84.182, 122.084, -177.849, 37.922, 178.303]
  MoveL 2343 to (-200, -42.4, 22.48) mm, rotated rx 90 ry 0 rz 180 deg; joints [1.351, -84.181, 122.083, -177.802, 37.922, 178.266]
  MoveL 2344 to (0, -42.4, 22.48) mm, rotated rx 90 ry 0 rz 180 deg; joints [1.154, -71.695, 106.629, -177.985, 34.951, 178.349]
  MoveL 2345 to (0, -42.4, 21.88) mm, rotated rx 90 ry 0 rz 180 deg; joints [1.179, -71.694, 106.628, -177.942, 34.951, 178.313]
  MoveL 2346 to (-200, -42.4, 21.88) mm, rotated rx 90 ry 0 rz 180 deg; joints [1.38, -84.18, 122.082, -177.754, 37.923, 178.228]
  MoveL 2347 to (-200, -42.4, 21.28) mm, rotated rx 90 ry 0 rz 180 deg; joints [1.409, -84.179, 122.081, -177.706, 37.924, 178.19]
  MoveL 2348 to (0, -42.4, 21.28) mm, rotated rx 90 ry 0 rz 180 deg; joints [1.204, -71.694, 106.627, -177.898, 34.952, 178.277]
  MoveL 2349 to (0, -42.4, 20.68) mm, rotated rx 90 ry 0 rz 180 deg; joints [1.229, -71.693, 106.626, -177.854, 34.952, 178.241]
  MoveL 2350 to (-200, -42.4, 20.68) mm, rotated rx 90 ry 0 rz 180 deg; joints [1.439, -84.178, 122.08, -177.659, 37.925, 178.153]
  MoveL 2351 to (-200, -42.4, 20.08) mm, rotated rx 90 ry 0 rz 180 deg; joints [1.468, -84.177, 122.079, -177.611, 37.926, 178.115]
  MoveL 2352 to (0, -42.4, 20.08) mm, rotated rx 90 ry 0 rz 180 deg; joints [1.254, -71.692, 106.625, -177.811, 34.953, 178.205]
  MoveL 2353 to (0, -42.4, 19.48) mm, rotated rx 90 ry 0 rz 180 deg; joints [1.279, -71.691, 106.624, -177.767, 34.953, 178.169]
  MoveL 2354 to (-200, -42.4, 19.48) mm, rotated rx 90 ry 0 rz 180 deg; joints [1.497, -84.176, 122.078, -177.563, 37.926, 178.078]
  MoveL 2355 to (-200, -42.4, 18.88) mm, rotated rx 90 ry 0 rz 180 deg; joints [1.527, -84.175, 122.076, -177.516, 37.927, 178.04]
  MoveL 2356 to (0, -42.4, 18.88) mm, rotated rx 90 ry 0 rz 180 deg; joints [1.304, -71.69, 106.623, -177.723, 34.954, 178.134]
  MoveL 2357 to (0, -42.4, 18.28) mm, rotated rx 90 ry 0 rz 180 deg; joints [1.329, -71.69, 106.622, -177.679, 34.954, 178.098]
  MoveL 2358 to (-200, -42.4, 18.28) mm, rotated rx 90 ry 0 rz 180 deg; joints [1.556, -84.174, 122.075, -177.468, 37.928, 178.002]
  MoveL 2359 to (-200, -42.4, 17.68) mm, rotated rx 90 ry 0 rz 180 deg; joints [1.585, -84.173, 122.074, -177.42, 37.929, 177.965]
  MoveL 2360 to (0, -42.4, 17.68) mm, rotated rx 90 ry 0 rz 180 deg; joints [1.354, -71.689, 106.621, -177.636, 34.955, 178.062]
  MoveL 2361 to (0, -42.4, 17.08) mm, rotated rx 90 ry 0 rz 180 deg; joints [1.379, -71.688, 106.619, -177.592, 34.955, 178.026]
  MoveL 2362 to (-200, -42.4, 17.08) mm, rotated rx 90 ry 0 rz 180 deg; joints [1.615, -84.172, 122.073, -177.373, 37.93, 177.927]
  MoveL 2363 to (-200, -42.4, 16.48) mm, rotated rx 90 ry 0 rz 180 deg; joints [1.644, -84.171, 122.072, -177.325, 37.931, 177.89]
  MoveL 2364 to (0, -42.4, 16.48) mm, rotated rx 90 ry 0 rz 180 deg; joints [1.404, -71.687, 106.618, -177.548, 34.956, 177.99]
  MoveL 2365 to (0, -42.4, 15.88) mm, rotated rx 90 ry 0 rz 180 deg; joints [1.429, -71.686, 106.617, -177.505, 34.957, 177.954]
  MoveL 2366 to (-200, -42.4, 15.88) mm, rotated rx 90 ry 0 rz 180 deg; joints [1.673, -84.17, 122.07, -177.277, 37.932, 177.852]
  MoveL 2367 to (-200, -42.4, 15.28) mm, rotated rx 90 ry 0 rz 180 deg; joints [1.703, -84.169, 122.069, -177.23, 37.933, 177.814]
  MoveL 2368 to (0, -42.4, 15.28) mm, rotated rx 90 ry 0 rz 180 deg; joints [1.454, -71.685, 106.616, -177.461, 34.957, 177.919]
  MoveL 2369 to (0, -42.4, 14.68) mm, rotated rx 88.51 ry 0 rz 180 deg; joints [1.868, -71.696, 106.555, -176.735, 34.903, 175.833]
  MoveL 2370 to (-200, -42.4, 14.68) mm, rotated rx 88.51 ry 0 rz 180 deg; joints [2.186, -84.181, 122.005, -176.438, 37.878, 175.699]
  MoveL 2371 to (-200, -42.37, 14.08) mm, rotated rx 85.74 ry 0 rz 180 deg; joints [3.064, -84.168, 121.898, -175.001, 37.836, 171.787]
  MoveL 2372 to (0, -42.37, 14.08) mm, rotated rx 85.74 ry 0 rz 180 deg; joints [2.618, -71.686, 106.452, -175.416, 34.851, 171.974]
  MoveL 2373 to (0, -42.31, 13.48) mm, rotated rx 82.97 ry 0 rz 180 deg; joints [3.368, -71.637, 106.361, -174.101, 34.866, 168.121]
  MoveL 2374 to (-200, -42.31, 13.48) mm, rotated rx 82.97 ry 0 rz 180 deg; joints [3.941, -84.108, 121.807, -173.571, 37.873, 167.884]
  MoveL 2375 to (-200, -42.22, 12.89) mm, rotated rx 80.19 ry 0 rz 180 deg; joints [4.817, -84.001, 121.73, -172.158, 37.989, 163.999]
  MoveL 2376 to (0, -42.22, 12.89) mm, rotated rx 80.19 ry 0 rz 180 deg; joints [4.118, -71.549, 106.284, -172.799, 34.947, 164.281]
  MoveL 2377 to (0, -42.1, 12.3) mm, rotated rx 77.42 ry 0 rz 180 deg; joints [4.863, -71.422, 106.219, -171.52, 35.093, 160.466]
  MoveL 2378 to (-200, -42.1, 12.3) mm, rotated rx 77.42 ry 0 rz 180 deg; joints [5.688, -83.847, 121.668, -170.773, 38.183, 160.145]
  MoveL 2379 to (-200, -41.96, 11.72) mm, rotated rx 74.65 ry 0 rz 180 deg; joints [6.552, -83.648, 121.621, -169.426, 38.451, 156.333]
  MoveL 2380 to (0, -41.96, 11.72) mm, rotated rx 74.65 ry 0 rz 180 deg; joints [5.604, -71.257, 106.168, -170.272, 35.302, 156.685]
  MoveL 2381 to (0, -41.78, 11.14) mm, rotated rx 71.88 ry 0 rz 180 deg; joints [6.337, -71.053, 106.129, -169.062, 35.572, 152.944]
  MoveL 2382 to (-200, -41.78, 11.14) mm, rotated rx 71.88 ry 0 rz 180 deg; joints [7.407, -83.402, 121.59, -168.124, 38.792, 152.569]
  MoveL 2383 to (-200, -41.59, 10.58) mm, rotated rx 69.11 ry 0 rz 180 deg; joints [8.251, -83.112, 121.573, -166.877, 39.202, 148.864]
  MoveL 2384 to (0, -41.59, 10.58) mm, rotated rx 69.11 ry 0 rz 180 deg; joints [7.061, -70.812, 106.104, -167.899, 35.902, 149.253]
  MoveL 2385 to (0, -41.36, 10.02) mm, rotated rx 66.33 ry 0 rz 180 deg; joints [7.774, -70.533, 106.091, -166.789, 36.288, 145.618]
  MoveL 2386 to (-200, -41.36, 10.02) mm, rotated rx 66.33 ry 0 rz 180 deg; joints [9.08, -82.777, 121.571, -165.69, 39.679, 145.226]
  MoveL 2387 to (-200, -41.1, 9.48) mm, rotated rx 63.56 ry 0 rz 180 deg; joints [9.894, -82.398, 121.583, -164.568, 40.218, 141.657]
  MoveL 2388 to (0, -41.1, 9.48) mm, rotated rx 63.56 ry 0 rz 180 deg; joints [8.474, -70.218, 106.091, -165.735, 36.729, 142.042]
  MoveL 2389 to (0, -40.82, 8.95) mm, rotated rx 60.79 ry 0 rz 180 deg; joints [9.159, -69.868, 106.103, -164.742, 37.22, 138.533]
  MoveL 2390 to (-200, -40.82, 8.95) mm, rotated rx 60.79 ry 0 rz 180 deg; joints [10.689, -81.977, 121.608, -163.515, 40.817, 138.164]
  MoveL 2391 to (-200, -40.52, 8.43) mm, rotated rx 58.01 ry 0 rz 180 deg; joints [11.465, -81.514, 121.647, -162.534, 41.471, 134.749]
  MoveL 2392 to (0, -40.52, 8.43) mm, rotated rx 58.01 ry 0 rz 180 deg; joints [9.829, -69.482, 106.127, -163.813, 37.76, 135.09]
  MoveL 2393 to (0, -40.19, 7.93) mm, rotated rx 55.24 ry 0 rz 180 deg; joints [10.48, -69.063, 106.162, -162.95, 38.345, 131.719]
  MoveL 2394 to (-200, -40.19, 7.93) mm, rotated rx 55.24 ry 0 rz 180 deg; joints [12.219, -81.01, 121.699, -161.625, 42.176, 131.414]
  MoveL 2395 to (-200, -39.83, 7.45) mm, rotated rx 52.47 ry 0 rz 180 deg; joints [12.95, -80.466, 121.763, -160.791, 42.929, 128.159]
  MoveL 2396 to (0, -39.83, 7.45) mm, rotated rx 52.47 ry 0 rz 180 deg; joints [11.113, -68.609, 106.208, -162.155, 38.972, 128.419]
  MoveL 2397 to (0, -39.46, 6.98) mm, rotated rx 49.7 ry 0 rz 180 deg; joints [11.724, -68.124, 106.264, -161.426, 39.638, 125.189]
  MoveL 2398 to (-200, -39.46, 6.98) mm, rotated rx 49.7 ry 0 rz 180 deg; joints [13.656, -79.884, 121.838, -160.029, 43.726, 124.984]
  MoveL 2399 to (-200, -39.06, 6.53) mm, rotated rx 46.93 ry 0 rz 180 deg; joints [14.335, -79.263, 121.924, -159.339, 44.563, 121.887]
  MoveL 2400 to (0, -39.06, 6.53) mm, rotated rx 46.93 ry 0 rz 180 deg; joints [12.314, -67.607, 106.33, -160.763, 40.339, 122.031]
  MoveL 2401 to (0, -38.64, 6.1) mm, rotated rx 44.15 ry 0 rz 180 deg; joints [12.881, -67.059, 106.405, -160.167, 41.073, 118.943]
  MoveL 2402 to (-200, -38.64, 6.1) mm, rotated rx 44.15 ry 0 rz 180 deg; joints [14.987, -78.606, 122.02, -158.719, 45.436, 118.867]
  MoveL 2403 to (-200, -38.2, 5.7) mm, rotated rx 41.38 ry 0 rz 180 deg; joints [15.609, -77.914, 122.125, -158.166, 46.344, 115.92]
  MoveL 2404 to (0, -38.2, 5.7) mm, rotated rx 41.38 ry 0 rz 180 deg; joints [13.423, -66.482, 106.489, -159.634, 41.838, 115.921]
  MoveL 2405 to (0, -37.74, 5.31) mm, rotated rx 38.61 ry 0 rz 180 deg; joints [13.94, -65.877, 106.581, -159.163, 42.629, 112.965]
  MoveL 2406 to (-200, -37.74, 5.31) mm, rotated rx 38.61 ry 0 rz 180 deg; joints [16.202, -77.187, 122.239, -157.679, 47.28, 113.045]
  MoveL 2407 to (-200, -37.26, 4.95) mm, rotated rx 35.84 ry 0 rz 180 deg; joints [16.764, -76.427, 122.36, -157.255, 48.245, 110.237]
  MoveL 2408 to (0, -37.26, 4.95) mm, rotated rx 35.84 ry 0 rz 180 deg; joints [14.43, -65.244, 106.68, -158.753, 43.444, 110.071]
  MoveL 2409 to (0, -36.77, 4.61) mm, rotated rx 33.06 ry 0 rz 180 deg; joints [14.893, -64.585, 106.785, -158.4, 44.282, 107.238]
  MoveL 2410 to (-200, -36.77, 4.61) mm, rotated rx 33.06 ry 0 rz 180 deg; joints [17.294, -75.637, 122.487, -156.89, 49.233, 107.493]
  MoveL 2411 to (-200, -36.26, 4.29) mm, rotated rx 30.29 ry 0 rz 180 deg; joints [17.791, -74.816, 122.621, -156.582, 50.242, 104.809]
  MoveL 2412 to (0, -36.26, 4.29) mm, rotated rx 30.29 ry 0 rz 180 deg; joints [15.329, -63.902, 106.896, -158.102, 45.138, 104.462]
  MoveL 2413 to (0, -35.73, 4) mm, rotated rx 27.52 ry 0 rz 180 deg; joints [15.735, -63.195, 107.013, -157.857, 46.012, 101.738]
  MoveL 2414 to (-200, -35.73, 4) mm, rotated rx 27.52 ry 0 rz 180 deg; joints [18.254, -73.966, 122.759, -156.327, 51.272, 102.181]
  MoveL 2415 to (-200, -35.19, 3.74) mm, rotated rx 24.75 ry 0 rz 180 deg; joints [18.683, -73.09, 122.902, -156.123, 52.317, 99.606]
  MoveL 2416 to (0, -35.19, 3.74) mm, rotated rx 24.75 ry 0 rz 180 deg; joints [16.112, -62.466, 107.133, -157.662, 46.901, 99.065]
  MoveL 2417 to (0, -34.64, 3.5) mm, rotated rx 21.98 ry 0 rz 180 deg; joints [16.459, -61.716, 107.258, -157.515, 47.803, 96.438]
  MoveL 2418 to (-200, -34.64, 3.5) mm, rotated rx 21.98 ry 0 rz 180 deg; joints [19.078, -72.188, 123.048, -155.967, 53.377, 97.079]
  MoveL 2419 to (-200, -34.08, 3.29) mm, rotated rx 19.2 ry 0 rz 180 deg; joints [19.438, -71.262, 123.196, -155.856, 54.45, 94.595]
  MoveL 2420 to (0, -34.08, 3.29) mm, rotated rx 19.2 ry 0 rz 180 deg; joints [16.776, -60.946, 107.385, -157.412, 48.715, 93.853]
  MoveL 2421 to (0, -33.51, 3.11) mm, rotated rx 16.43 ry 0 rz 180 deg; joints [17.061, -60.159, 107.515, -157.353, 49.637, 91.31]
  MoveL 2422 to (-200, -33.51, 3.11) mm, rotated rx 16.43 ry 0 rz 180 deg; joints [19.762, -70.314, 123.347, -155.788, 55.532, 92.152]
  MoveL 2423 to (-200, -32.93, 2.95) mm, rotated rx 13.66 ry 0 rz 180 deg; joints [20.05, -69.345, 123.498, -155.761, 56.624, 89.745]
  MoveL 2424 to (0, -32.93, 2.95) mm, rotated rx 13.66 ry 0 rz 180 deg; joints [17.315, -59.355, 107.647, -157.335, 50.566, 88.801]
  MoveL 2425 to (0, -32.34, 2.82) mm, rotated rx 10.88 ry 0 rz 180 deg; joints [17.538, -58.536, 107.779, -157.354, 51.5, 86.326]
  MoveL 2426 to (-200, -32.34, 2.82) mm, rotated rx 10.88 ry 0 rz 180 deg; joints [20.302, -68.358, 123.65, -155.771, 57.722, 87.372]
  MoveL 2427 to (-200, -31.75, 2.72) mm, rotated rx 8.11 ry 0 rz 180 deg; joints [20.517, -67.354, 123.801, -155.817, 58.825, 85.027]
  MoveL 2428 to (0, -31.75, 2.72) mm, rotated rx 8.11 ry 0 rz 180 deg; joints [17.728, -57.705, 107.913, -157.411, 52.439, 83.882]
  MoveL 2429 to (0, -31.15, 2.65) mm, rotated rx 5.34 ry 0 rz 180 deg; joints [17.886, -56.861, 108.046, -157.502, 53.38, 81.462]
  MoveL 2430 to (-200, -31.15, 2.65) mm, rotated rx 5.34 ry 0 rz 180 deg; joints [20.696, -66.335, 123.952, -155.898, 59.933, 82.707]
  MoveL 2431 to (-200, -30.56, 2.61) mm, rotated rx 2.57 ry 0 rz 180 deg; joints [20.838, -65.303, 124.101, -156.011, 61.042, 80.409]
  MoveL 2432 to (0, -30.56, 2.61) mm, rotated rx 2.57 ry 0 rz 180 deg; joints [18.011, -56.007, 108.179, -157.626, 54.321, 79.068]
  MoveL 2433 to (0, -29.96, 2.6) mm, rotated rx 0 ry 0 rz 180 deg; joints [18.098, -55.207, 108.302, -157.77, 55.195, 76.869]
  MoveL 2434 to (-200, -29.96, 2.6) mm, rotated rx 0 ry 0 rz 180 deg; joints [20.936, -64.334, 124.237, -156.144, 62.072, 78.299]
  MoveL 2435 to (-200, -29.36, 2.6) mm, rotated rx 0 ry 0 rz 180 deg; joints [20.936, -64.3, 124.244, -156.153, 62.109, 78.317]
  MoveL 2436 to (0, -29.36, 2.6) mm, rotated rx 0 ry 0 rz 180 deg; joints [18.098, -55.179, 108.308, -157.779, 55.227, 76.884]
  MoveL 2437 to (0, -28.76, 2.6) mm, rotated rx 0 ry 0 rz 180 deg; joints [18.098, -55.151, 108.315, -157.788, 55.259, 76.9]
  MoveL 2438 to (-200, -28.76, 2.6) mm, rotated rx 0 ry 0 rz 180 deg; joints [20.936, -64.266, 124.251, -156.162, 62.147, 78.336]
  MoveL 2439 to (-200, -28.16, 2.6) mm, rotated rx 0 ry 0 rz 180 deg; joints [20.936, -64.233, 124.258, -156.17, 62.184, 78.355]
  MoveL 2440 to (0, -28.16, 2.6) mm, rotated rx 0 ry 0 rz 180 deg; joints [18.098, -55.123, 108.321, -157.797, 55.291, 76.916]
  MoveL 2441 to (0, -27.56, 2.6) mm, rotated rx 0 ry 0 rz 180 deg; joints [18.098, -55.095, 108.327, -157.806, 55.322, 76.932]
  MoveL 2442 to (-200, -27.56, 2.6) mm, rotated rx 0 ry 0 rz 180 deg; joints [20.936, -64.199, 124.264, -156.179, 62.221, 78.373]
  MoveL 2443 to (-200, -26.96, 2.6) mm, rotated rx 0 ry 0 rz 180 deg; joints [20.936, -64.165, 124.271, -156.188, 62.259, 78.392]
  MoveL 2444 to (0, -26.96, 2.6) mm, rotated rx 0 ry 0 rz 180 deg; joints [18.098, -55.067, 108.333, -157.814, 55.354, 76.947]
  MoveL 2445 to (0, -26.36, 2.6) mm, rotated rx 0 ry 0 rz 180 deg; joints [18.098, -55.039, 108.339, -157.823, 55.386, 76.963]
  MoveL 2446 to (-200, -26.36, 2.6) mm, rotated rx 0 ry 0 rz 180 deg; joints [20.936, -64.131, 124.278, -156.196, 62.296, 78.41]
  MoveL 2447 to (-200, -25.76, 2.6) mm, rotated rx 0 ry 0 rz 180 deg; joints [20.936, -64.096, 124.285, -156.205, 62.333, 78.429]
  MoveL 2448 to (0, -25.76, 2.6) mm, rotated rx 0 ry 0 rz 180 deg; joints [18.098, -55.011, 108.346, -157.832, 55.417, 76.979]
  MoveL 2449 to (0, -25.16, 2.6) mm, rotated rx 0 ry 0 rz 180 deg; joints [18.098, -54.983, 108.352, -157.841, 55.449, 76.994]
  MoveL 2450 to (-200, -25.16, 2.6) mm, rotated rx 0 ry 0 rz 180 deg; joints [20.936, -64.062, 124.291, -156.214, 62.37, 78.447]
  MoveL 2451 to (-200, -24.56, 2.6) mm, rotated rx 0 ry 0 rz 180 deg; joints [20.936, -64.028, 124.298, -156.222, 62.408, 78.466]
  MoveL 2452 to (0, -24.56, 2.6) mm, rotated rx 0 ry 0 rz 180 deg; joints [18.098, -54.955, 108.358, -157.85, 55.481, 77.01]
  MoveL 2453 to (0, -23.96, 2.6) mm, rotated rx 0 ry 0 rz 180 deg; joints [18.098, -54.927, 108.364, -157.859, 55.512, 77.026]
  MoveL 2454 to (-200, -23.96, 2.6) mm, rotated rx 0 ry 0 rz 180 deg; joints [20.936, -63.994, 124.304, -156.231, 62.445, 78.485]
  MoveL 2455 to (-200, -23.36, 2.6) mm, rotated rx 0 ry 0 rz 180 deg; joints [20.936, -63.96, 124.311, -156.239, 62.482, 78.503]
  MoveL 2456 to (0, -23.36, 2.6) mm, rotated rx 0 ry 0 rz 180 deg; joints [18.098, -54.899, 108.37, -157.868, 55.544, 77.041]
  MoveL 2457 to (0, -22.76, 2.6) mm, rotated rx 0 ry 0 rz 180 deg; joints [18.098, -54.871, 108.376, -157.877, 55.575, 77.057]
  MoveL 2458 to (-200, -22.76, 2.6) mm, rotated rx 0 ry 0 rz 180 deg; joints [20.936, -63.926, 124.318, -156.248, 62.519, 78.521]
  MoveL 2459 to (-200, -22.16, 2.6) mm, rotated rx 0 ry 0 rz 180 deg; joints [20.936, -63.892, 124.324, -156.256, 62.557, 78.54]
  MoveL 2460 to (0, -22.16, 2.6) mm, rotated rx 0 ry 0 rz 180 deg; joints [18.098, -54.842, 108.382, -157.885, 55.607, 77.072]
  MoveL 2461 to (0, -21.56, 2.6) mm, rotated rx 0 ry 0 rz 180 deg; joints [18.098, -54.814, 108.388, -157.894, 55.639, 77.088]
  MoveL 2462 to (-200, -21.56, 2.6) mm, rotated rx 0 ry 0 rz 180 deg; joints [20.936, -63.857, 124.331, -156.265, 62.594, 78.558]
  MoveL 2463 to (-200, -20.96, 2.6) mm, rotated rx 0 ry 0 rz 180 deg; joints [20.936, -63.823, 124.337, -156.273, 62.631, 78.577]
  MoveL 2464 to (0, -20.96, 2.6) mm, rotated rx 0 ry 0 rz 180 deg; joints [18.098, -54.786, 108.394, -157.903, 55.67, 77.104]
  MoveL 2465 to (0, -20.36, 2.6) mm, rotated rx 0 ry 0 rz 180 deg; joints [18.098, -54.758, 108.4, -157.912, 55.702, 77.119]
  MoveL 2466 to (-200, -20.36, 2.6) mm, rotated rx 0 ry 0 rz 180 deg; joints [20.936, -63.789, 124.343, -156.282, 62.668, 78.595]
  MoveL 2467 to (-200, -19.76, 2.6) mm, rotated rx 0 ry 0 rz 180 deg; joints [20.936, -63.755, 124.35, -156.29, 62.706, 78.614]
  MoveL 2468 to (0, -19.76, 2.6) mm, rotated rx 0 ry 0 rz 180 deg; joints [18.098, -54.73, 108.406, -157.92, 55.733, 77.135]
  MoveL 2469 to (0, -19.16, 2.6) mm, rotated rx 0 ry 0 rz 180 deg; joints [18.098, -54.701, 108.411, -157.929, 55.765, 77.15]
  MoveL 2470 to (-200, -19.16, 2.6) mm, rotated rx 0 ry 0 rz 180 deg; joints [20.936, -63.72, 124.356, -156.299, 62.743, 78.632]
  MoveL 2471 to (-200, -18.56, 2.6) mm, rotated rx 0 ry 0 rz 180 deg; joints [20.936, -63.686, 124.362, -156.307, 62.78, 78.65]
  MoveL 2472 to (0, -18.56, 2.6) mm, rotated rx 0 ry 0 rz 180 deg; joints [18.098, -54.673, 108.417, -157.938, 55.796, 77.166]
  MoveL 2473 to (0, -17.96, 2.6) mm, rotated rx 0 ry 0 rz 180 deg; joints [18.098, -54.645, 108.423, -157.946, 55.828, 77.181]
  MoveL 2474 to (-200, -17.96, 2.6) mm, rotated rx 0 ry 0 rz 180 deg; joints [20.936, -63.652, 124.369, -156.316, 62.817, 78.669]
  MoveL 2475 to (-200, -17.36, 2.6) mm, rotated rx 0 ry 0 rz 180 deg; joints [20.936, -63.617, 124.375, -156.324, 62.854, 78.687]
  MoveL 2476 to (0, -17.36, 2.6) mm, rotated rx 0 ry 0 rz 180 deg; joints [18.098, -54.617, 108.429, -157.955, 55.86, 77.196]
  MoveL 2477 to (0, -16.76, 2.6) mm, rotated rx 0 ry 0 rz 180 deg; joints [18.098, -54.588, 108.434, -157.964, 55.891, 77.212]
  MoveL 2478 to (-200, -16.76, 2.6) mm, rotated rx 0 ry 0 rz 180 deg; joints [20.936, -63.583, 124.381, -156.332, 62.891, 78.705]
  MoveL 2479 to (-200, -16.16, 2.6) mm, rotated rx 0 ry 0 rz 180 deg; joints [20.936, -63.549, 124.387, -156.341, 62.929, 78.724]
  MoveL 2480 to (0, -16.16, 2.6) mm, rotated rx 0 ry 0 rz 180 deg; joints [18.098, -54.56, 108.44, -157.972, 55.923, 77.227]
  MoveL 2481 to (0, -15.56, 2.6) mm, rotated rx 0 ry 0 rz 180 deg; joints [18.098, -54.532, 108.446, -157.981, 55.954, 77.243]
  MoveL 2482 to (-200, -15.56, 2.6) mm, rotated rx 0 ry 0 rz 180 deg; joints [20.936, -63.514, 124.393, -156.349, 62.966, 78.742]
  MoveL 2483 to (-200, -14.96, 2.6) mm, rotated rx 0 ry 0 rz 180 deg; joints [20.936, -63.48, 124.4, -156.357, 63.003, 78.76]
  MoveL 2484 to (0, -14.96, 2.6) mm, rotated rx 0 ry 0 rz 180 deg; joints [18.098, -54.503, 108.451, -157.99, 55.986, 77.258]
  MoveL 2485 to (0, -14.36, 2.6) mm, rotated rx 0 ry 0 rz 180 deg; joints [18.098, -54.475, 108.457, -157.998, 56.017, 77.273]
  MoveL 2486 to (-200, -14.36, 2.6) mm, rotated rx 0 ry 0 rz 180 deg; joints [20.936, -63.445, 124.406, -156.365, 63.04, 78.778]
  MoveL 2487 to (-200, -13.76, 2.6) mm, rotated rx 0 ry 0 rz 180 deg; joints [20.936, -63.411, 124.412, -156.374, 63.077, 78.797]
  MoveL 2488 to (0, -13.76, 2.6) mm, rotated rx 0 ry 0 rz 180 deg; joints [18.098, -54.447, 108.463, -158.007, 56.049, 77.289]
  MoveL 2489 to (0, -13.16, 2.6) mm, rotated rx 0 ry 0 rz 180 deg; joints [18.098, -54.418, 108.468, -158.015, 56.08, 77.304]
  MoveL 2490 to (-200, -13.16, 2.6) mm, rotated rx 0 ry 0 rz 180 deg; joints [20.936, -63.376, 124.418, -156.382, 63.114, 78.815]
  MoveL 2491 to (-200, -12.56, 2.6) mm, rotated rx 0 ry 0 rz 180 deg; joints [20.936, -63.342, 124.424, -156.39, 63.151, 78.833]
  MoveL 2492 to (0, -12.56, 2.6) mm, rotated rx 0 ry 0 rz 180 deg; joints [18.098, -54.39, 108.474, -158.024, 56.112, 77.319]
  MoveL 2493 to (0, -11.96, 2.6) mm, rotated rx 0 ry 0 rz 180 deg; joints [18.098, -54.361, 108.479, -158.032, 56.143, 77.335]
  MoveL 2494 to (-200, -11.96, 2.6) mm, rotated rx 0 ry 0 rz 180 deg; joints [20.936, -63.307, 124.43, -156.398, 63.189, 78.851]
  MoveL 2495 to (-200, -11.36, 2.6) mm, rotated rx 0 ry 0 rz 180 deg; joints [20.936, -63.273, 124.436, -156.407, 63.226, 78.869]
  MoveL 2496 to (0, -11.36, 2.6) mm, rotated rx 0 ry 0 rz 180 deg; joints [18.098, -54.333, 108.485, -158.041, 56.175, 77.35]
  MoveL 2497 to (0, -10.76, 2.6) mm, rotated rx 0 ry 0 rz 180 deg; joints [18.098, -54.304, 108.49, -158.049, 56.206, 77.365]
  MoveL 2498 to (-200, -10.76, 2.6) mm, rotated rx 0 ry 0 rz 180 deg; joints [20.936, -63.238, 124.441, -156.415, 63.263, 78.888]
  MoveL 2499 to (-200, -10.16, 2.6) mm, rotated rx 0 ry 0 rz 180 deg; joints [20.936, -63.203, 124.447, -156.423, 63.3, 78.906]
  MoveL 2500 to (0, -10.16, 2.6) mm, rotated rx 0 ry 0 rz 180 deg; joints [18.098, -54.276, 108.495, -158.058, 56.237, 77.38]
  MoveL 2501 to (0, -9.56, 2.6) mm, rotated rx 0 ry 0 rz 180 deg; joints [18.098, -54.247, 108.501, -158.066, 56.269, 77.396]
  MoveL 2502 to (-200, -9.56, 2.6) mm, rotated rx 0 ry 0 rz 180 deg; joints [20.936, -63.169, 124.453, -156.431, 63.337, 78.924]
  MoveL 2503 to (-200, -8.96, 2.6) mm, rotated rx 0 ry 0 rz 180 deg; joints [20.936, -63.134, 124.459, -156.439, 63.374, 78.942]
  MoveL 2504 to (0, -8.96, 2.6) mm, rotated rx 0 ry 0 rz 180 deg; joints [18.098, -54.219, 108.506, -158.075, 56.3, 77.411]
  MoveL 2505 to (0, -8.36, 2.6) mm, rotated rx 0 ry 0 rz 180 deg; joints [18.098, -54.19, 108.511, -158.083, 56.332, 77.426]
  MoveL 2506 to (-200, -8.36, 2.6) mm, rotated rx 0 ry 0 rz 180 deg; joints [20.936, -63.1, 124.465, -156.447, 63.411, 78.96]
  MoveL 2507 to (-200, -7.76, 2.6) mm, rotated rx 0 ry 0 rz 180 deg; joints [20.936, -63.065, 124.47, -156.455, 63.448, 78.978]
  MoveL 2508 to (0, -7.76, 2.6) mm, rotated rx 0 ry 0 rz 180 deg; joints [18.098, -54.162, 108.517, -158.092, 56.363, 77.441]
  MoveL 2509 to (0, -7.16, 2.6) mm, rotated rx 0 ry 0 rz 180 deg; joints [18.098, -54.133, 108.522, -158.1, 56.394, 77.456]
  MoveL 2510 to (-200, -7.16, 2.6) mm, rotated rx 0 ry 0 rz 180 deg; joints [20.936, -63.03, 124.476, -156.463, 63.485, 78.996]
  MoveL 2511 to (-200, -6.56, 2.6) mm, rotated rx 0 ry 0 rz 180 deg; joints [20.936, -62.995, 124.482, -156.471, 63.522, 79.014]
  MoveL 2512 to (0, -6.56, 2.6) mm, rotated rx 0 ry 0 rz 180 deg; joints [18.098, -54.105, 108.527, -158.108, 56.426, 77.471]
  MoveL 2513 to (0, -5.96, 2.6) mm, rotated rx 0 ry 0 rz 180 deg; joints [18.098, -54.076, 108.532, -158.117, 56.457, 77.487]
  MoveL 2514 to (-200, -5.96, 2.6) mm, rotated rx 0 ry 0 rz 180 deg; joints [20.936, -62.961, 124.487, -156.479, 63.559, 79.032]
  MoveL 2515 to (-200, -5.36, 2.6) mm, rotated rx 0 ry 0 rz 180 deg; joints [20.936, -62.926, 124.493, -156.487, 63.596, 79.05]
  MoveL 2516 to (0, -5.36, 2.6) mm, rotated rx 0 ry 0 rz 180 deg; joints [18.098, -54.047, 108.538, -158.125, 56.489, 77.502]
  MoveL 2517 to (0, -4.76, 2.6) mm, rotated rx 0 ry 0 rz 180 deg; joints [18.098, -54.019, 108.543, -158.133, 56.52, 77.517]
  MoveL 2518 to (-200, -4.76, 2.6) mm, rotated rx 0 ry 0 rz 180 deg; joints [20.936, -62.891, 124.499, -156.495, 63.633, 79.068]
  MoveL 2519 to (-200, -4.16, 2.6) mm, rotated rx 0 ry 0 rz 180 deg; joints [20.936, -62.856, 124.504, -156.503, 63.67, 79.086]
  MoveL 2520 to (0, -4.16, 2.6) mm, rotated rx 0 ry 0 rz 180 deg; joints [18.098, -53.99, 108.548, -158.142, 56.551, 77.532]
  MoveL 2521 to (0, -3.56, 2.6) mm, rotated rx 0 ry 0 rz 180 deg; joints [18.098, -53.961, 108.553, -158.15, 56.583, 77.547]
  MoveL 2522 to (-200, -3.56, 2.6) mm, rotated rx 0 ry 0 rz 180 deg; joints [20.936, -62.821, 124.51, -156.511, 63.707, 79.104]
  MoveL 2523 to (-200, -2.96, 2.6) mm, rotated rx 0 ry 0 rz 180 deg; joints [20.936, -62.786, 124.515, -156.519, 63.744, 79.122]
  MoveL 2524 to (0, -2.96, 2.6) mm, rotated rx 0 ry 0 rz 180 deg; joints [18.098, -53.933, 108.558, -158.158, 56.614, 77.562]
  MoveL 2525 to (0, -2.36, 2.6) mm, rotated rx 0 ry 0 rz 180 deg; joints [18.098, -53.904, 108.563, -158.167, 56.645, 77.577]
  MoveL 2526 to (-200, -2.36, 2.6) mm, rotated rx 0 ry 0 rz 180 deg; joints [20.936, -62.752, 124.521, -156.527, 63.781, 79.14]
  MoveL 2527 to (-200, -1.76, 2.6) mm, rotated rx 0 ry 0 rz 180 deg; joints [20.936, -62.717, 124.526, -156.535, 63.818, 79.158]
  MoveL 2528 to (0, -1.76, 2.6) mm, rotated rx 0 ry 0 rz 180 deg; joints [18.098, -53.875, 108.568, -158.175, 56.677, 77.592]
  MoveL 2529 to (0, -1.16, 2.6) mm, rotated rx 0 ry 0 rz 180 deg; joints [18.098, -53.846, 108.573, -158.183, 56.708, 77.607]
  MoveL 2530 to (-200, -1.16, 2.6) mm, rotated rx 0 ry 0 rz 180 deg; joints [20.936, -62.682, 124.531, -156.543, 63.855, 79.176]
  MoveL 2531 to (-200, -0.56, 2.6) mm, rotated rx 0 ry 0 rz 180 deg; joints [20.936, -62.647, 124.537, -156.551, 63.892, 79.193]
  MoveL 2532 to (0, -0.56, 2.6) mm, rotated rx 0 ry 0 rz 180 deg; joints [18.098, -53.818, 108.578, -158.191, 56.739, 77.622]
  MoveL 2533 to (0, 0, 2.6) mm, rotated rx 0 ry 0 rz 180 deg; joints [18.098, -53.791, 108.582, -158.199, 56.768, 77.636]
  MoveL 2534 to (-200, 0, 2.6) mm, rotated rx 0 ry 0 rz 180 deg; joints [20.936, -62.614, 124.542, -156.558, 63.927, 79.21]
  MoveL 2535 to (-200, 0, 2.2) mm, rotated rx 0 ry 0 rz 180 deg; joints [20.954, -62.608, 124.53, -156.539, 63.925, 79.2]
  MoveL 2536 to (0, 0, 2.2) mm, rotated rx 0 ry 0 rz 180 deg; joints [18.113, -53.785, 108.571, -158.18, 56.767, 77.624]
  MoveL 2537 to (0, -0.6, 2.2) mm, rotated rx 0 ry 0 rz 180 deg; joints [18.113, -53.814, 108.566, -158.172, 56.735, 77.609]
  MoveL 2538 to (-200, -0.6, 2.2) mm, rotated rx 0 ry 0 rz 180 deg; joints [20.954, -62.643, 124.525, -156.531, 63.888, 79.182]
  MoveL 2539 to (-200, -1.2, 2.2) mm, rotated rx 0 ry 0 rz 180 deg; joints [20.954, -62.678, 124.52, -156.523, 63.851, 79.164]
  MoveL 2540 to (0, -1.2, 2.2) mm, rotated rx 0 ry 0 rz 180 deg; joints [18.113, -53.842, 108.561, -158.164, 56.704, 77.594]
  MoveL 2541 to (0, -1.8, 2.2) mm, rotated rx 0 ry 0 rz 180 deg; joints [18.113, -53.871, 108.556, -158.155, 56.673, 77.579]
  MoveL 2542 to (-200, -1.8, 2.2) mm, rotated rx 0 ry 0 rz 180 deg; joints [20.954, -62.713, 124.514, -156.515, 63.814, 79.146]
  MoveL 2543 to (-200, -2.4, 2.2) mm, rotated rx 0 ry 0 rz 180 deg; joints [20.954, -62.748, 124.509, -156.507, 63.777, 79.128]
  MoveL 2544 to (0, -2.4, 2.2) mm, rotated rx 0 ry 0 rz 180 deg; joints [18.113, -53.9, 108.551, -158.147, 56.641, 77.564]
  MoveL 2545 to (0, -3, 2.2) mm, rotated rx 0 ry 0 rz 180 deg; joints [18.113, -53.929, 108.546, -158.139, 56.61, 77.549]
  MoveL 2546 to (-200, -3, 2.2) mm, rotated rx 0 ry 0 rz 180 deg; joints [20.954, -62.782, 124.503, -156.499, 63.74, 79.11]
  MoveL 2547 to (-200, -3.6, 2.2) mm, rotated rx 0 ry 0 rz 180 deg; joints [20.954, -62.817, 124.498, -156.491, 63.703, 79.092]
  MoveL 2548 to (0, -3.6, 2.2) mm, rotated rx 0 ry 0 rz 180 deg; joints [18.113, -53.957, 108.541, -158.13, 56.579, 77.534]
  MoveL 2549 to (0, -4.2, 2.2) mm, rotated rx 0 ry 0 rz 180 deg; joints [18.113, -53.986, 108.536, -158.122, 56.547, 77.519]
  MoveL 2550 to (-200, -4.2, 2.2) mm, rotated rx 0 ry 0 rz 180 deg; joints [20.954, -62.852, 124.492, -156.483, 63.666, 79.074]
  MoveL 2551 to (-200, -4.8, 2.2) mm, rotated rx 0 ry 0 rz 180 deg; joints [20.954, -62.887, 124.487, -156.475, 63.629, 79.056]
  MoveL 2552 to (0, -4.8, 2.2) mm, rotated rx 0 ry 0 rz 180 deg; joints [18.113, -54.015, 108.531, -158.114, 56.516, 77.504]
  MoveL 2553 to (0, -5.4, 2.2) mm, rotated rx 0 ry 0 rz 180 deg; joints [18.113, -54.043, 108.526, -158.106, 56.485, 77.489]
  MoveL 2554 to (-200, -5.4, 2.2) mm, rotated rx 0 ry 0 rz 180 deg; joints [20.954, -62.922, 124.481, -156.467, 63.592, 79.038]
  MoveL 2555 to (-200, -6, 2.2) mm, rotated rx 0 ry 0 rz 180 deg; joints [20.954, -62.957, 124.476, -156.459, 63.555, 79.02]
  MoveL 2556 to (0, -6, 2.2) mm, rotated rx 0 ry 0 rz 180 deg; joints [18.113, -54.072, 108.521, -158.097, 56.453, 77.473]
  MoveL 2557 to (0, -6.6, 2.2) mm, rotated rx 0 ry 0 rz 180 deg; joints [18.113, -54.101, 108.516, -158.089, 56.422, 77.458]
  MoveL 2558 to (-200, -6.6, 2.2) mm, rotated rx 0 ry 0 rz 180 deg; joints [20.954, -62.991, 124.47, -156.451, 63.518, 79.002]
  MoveL 2559 to (-200, -7.2, 2.2) mm, rotated rx 0 ry 0 rz 180 deg; joints [20.954, -63.026, 124.464, -156.443, 63.481, 78.984]
  MoveL 2560 to (0, -7.2, 2.2) mm, rotated rx 0 ry 0 rz 180 deg; joints [18.113, -54.129, 108.511, -158.08, 56.391, 77.443]
  MoveL 2561 to (0, -7.8, 2.2) mm, rotated rx 0 ry 0 rz 180 deg; joints [18.113, -54.158, 108.505, -158.072, 56.359, 77.428]
  MoveL 2562 to (-200, -7.8, 2.2) mm, rotated rx 0 ry 0 rz 180 deg; joints [20.954, -63.061, 124.459, -156.435, 63.444, 78.966]
  MoveL 2563 to (-200, -8.4, 2.2) mm, rotated rx 0 ry 0 rz 180 deg; joints [20.954, -63.095, 124.453, -156.427, 63.407, 78.948]
  MoveL 2564 to (0, -8.4, 2.2) mm, rotated rx 0 ry 0 rz 180 deg; joints [18.113, -54.186, 108.5, -158.064, 56.328, 77.413]
  MoveL 2565 to (0, -9, 2.2) mm, rotated rx 0 ry 0 rz 180 deg; joints [18.113, -54.215, 108.495, -158.055, 56.297, 77.398]
  MoveL 2566 to (-200, -9, 2.2) mm, rotated rx 0 ry 0 rz 180 deg; joints [20.954, -63.13, 124.447, -156.419, 63.37, 78.93]
  MoveL 2567 to (-200, -9.6, 2.2) mm, rotated rx 0 ry 0 rz 180 deg; joints [20.954, -63.165, 124.441, -156.411, 63.333, 78.912]
  MoveL 2568 to (0, -9.6, 2.2) mm, rotated rx 0 ry 0 rz 180 deg; joints [18.113, -54.243, 108.489, -158.047, 56.265, 77.382]
  MoveL 2569 to (0, -10.2, 2.2) mm, rotated rx 0 ry 0 rz 180 deg; joints [18.113, -54.272, 108.484, -158.038, 56.234, 77.367]
  MoveL 2570 to (-200, -10.2, 2.2) mm, rotated rx 0 ry 0 rz 180 deg; joints [20.954, -63.199, 124.435, -156.403, 63.296, 78.894]
  MoveL 2571 to (-200, -10.8, 2.2) mm, rotated rx 0 ry 0 rz 180 deg; joints [20.954, -63.234, 124.43, -156.394, 63.259, 78.876]
  MoveL 2572 to (0, -10.8, 2.2) mm, rotated rx 0 ry 0 rz 180 deg; joints [18.113, -54.3, 108.479, -158.03, 56.202, 77.352]
  MoveL 2573 to (0, -11.4, 2.2) mm, rotated rx 0 ry 0 rz 180 deg; joints [18.113, -54.329, 108.473, -158.021, 56.171, 77.337]
  MoveL 2574 to (-200, -11.4, 2.2) mm, rotated rx 0 ry 0 rz 180 deg; joints [20.954, -63.269, 124.424, -156.386, 63.222, 78.857]
  MoveL 2575 to (-200, -12, 2.2) mm, rotated rx 0 ry 0 rz 180 deg; joints [20.954, -63.303, 124.418, -156.378, 63.185, 78.839]
  MoveL 2576 to (0, -12, 2.2) mm, rotated rx 0 ry 0 rz 180 deg; joints [18.113, -54.357, 108.468, -158.013, 56.139, 77.321]
  MoveL 2577 to (0, -12.6, 2.2) mm, rotated rx 0 ry 0 rz 180 deg; joints [18.113, -54.386, 108.462, -158.004, 56.108, 77.306]
  MoveL 2578 to (-200, -12.6, 2.2) mm, rotated rx 0 ry 0 rz 180 deg; joints [20.954, -63.338, 124.412, -156.37, 63.148, 78.821]
  MoveL 2579 to (-200, -13.2, 2.2) mm, rotated rx 0 ry 0 rz 180 deg; joints [20.954, -63.372, 124.406, -156.362, 63.11, 78.803]
  MoveL 2580 to (0, -13.2, 2.2) mm, rotated rx 0 ry 0 rz 180 deg; joints [18.113, -54.414, 108.457, -157.996, 56.076, 77.291]
  MoveL 2581 to (0, -13.8, 2.2) mm, rotated rx 0 ry 0 rz 180 deg; joints [18.113, -54.443, 108.451, -157.987, 56.045, 77.275]
  MoveL 2582 to (-200, -13.8, 2.2) mm, rotated rx 0 ry 0 rz 180 deg; joints [20.954, -63.407, 124.4, -156.353, 63.073, 78.785]
  MoveL 2583 to (-200, -14.4, 2.2) mm, rotated rx 0 ry 0 rz 180 deg; joints [20.954, -63.441, 124.394, -156.345, 63.036, 78.766]
  MoveL 2584 to (0, -14.4, 2.2) mm, rotated rx 0 ry 0 rz 180 deg; joints [18.113, -54.471, 108.446, -157.979, 56.014, 77.26]
  MoveL 2585 to (0, -15, 2.2) mm, rotated rx 0 ry 0 rz 180 deg; joints [18.113, -54.499, 108.44, -157.97, 55.982, 77.245]
  MoveL 2586 to (-200, -15, 2.2) mm, rotated rx 0 ry 0 rz 180 deg; joints [20.954, -63.476, 124.388, -156.337, 62.999, 78.748]
  MoveL 2587 to (-200, -15.6, 2.2) mm, rotated rx 0 ry 0 rz 180 deg; joints [20.954, -63.51, 124.381, -156.329, 62.962, 78.73]
  MoveL 2588 to (0, -15.6, 2.2) mm, rotated rx 0 ry 0 rz 180 deg; joints [18.113, -54.528, 108.434, -157.961, 55.951, 77.229]
  MoveL 2589 to (0, -16.2, 2.2) mm, rotated rx 0 ry 0 rz 180 deg; joints [18.113, -54.556, 108.429, -157.953, 55.919, 77.214]
  MoveL 2590 to (-200, -16.2, 2.2) mm, rotated rx 0 ry 0 rz 180 deg; joints [20.954, -63.545, 124.375, -156.32, 62.925, 78.712]
  MoveL 2591 to (-200, -16.8, 2.2) mm, rotated rx 0 ry 0 rz 180 deg; joints [20.954, -63.579, 124.369, -156.312, 62.888, 78.693]
  MoveL 2592 to (0, -16.8, 2.2) mm, rotated rx 0 ry 0 rz 180 deg; joints [18.113, -54.584, 108.423, -157.944, 55.888, 77.198]
  MoveL 2593 to (0, -17.4, 2.2) mm, rotated rx 0 ry 0 rz 180 deg; joints [18.113, -54.613, 108.417, -157.935, 55.856, 77.183]
  MoveL 2594 to (-200, -17.4, 2.2) mm, rotated rx 0 ry 0 rz 180 deg; joints [20.954, -63.613, 124.363, -156.304, 62.85, 78.675]
  MoveL 2595 to (-200, -18, 2.2) mm, rotated rx 0 ry 0 rz 180 deg; joints [20.954, -63.648, 124.357, -156.295, 62.813, 78.657]
  MoveL 2596 to (0, -18, 2.2) mm, rotated rx 0 ry 0 rz 180 deg; joints [18.113, -54.641, 108.411, -157.927, 55.824, 77.168]
  MoveL 2597 to (0, -18.6, 2.2) mm, rotated rx 0 ry 0 rz 180 deg; joints [18.113, -54.669, 108.406, -157.918, 55.793, 77.152]
  MoveL 2598 to (-200, -18.6, 2.2) mm, rotated rx 0 ry 0 rz 180 deg; joints [20.954, -63.682, 124.35, -156.287, 62.776, 78.638]
  MoveL 2599 to (-200, -19.2, 2.2) mm, rotated rx 0 ry 0 rz 180 deg; joints [20.954, -63.716, 124.344, -156.278, 62.739, 78.62]
  MoveL 2600 to (0, -19.2, 2.2) mm, rotated rx 0 ry 0 rz 180 deg; joints [18.113, -54.697, 108.4, -157.909, 55.761, 77.137]
  MoveL 2601 to (0, -19.8, 2.2) mm, rotated rx 0 ry 0 rz 180 deg; joints [18.113, -54.726, 108.394, -157.901, 55.73, 77.121]
  MoveL 2602 to (-200, -19.8, 2.2) mm, rotated rx 0 ry 0 rz 180 deg; joints [20.954, -63.751, 124.338, -156.27, 62.702, 78.601]
  MoveL 2603 to (-200, -20.4, 2.2) mm, rotated rx 0 ry 0 rz 180 deg; joints [20.954, -63.785, 124.331, -156.261, 62.665, 78.583]
  MoveL 2604 to (0, -20.4, 2.2) mm, rotated rx 0 ry 0 rz 180 deg; joints [18.113, -54.754, 108.388, -157.892, 55.698, 77.106]
  MoveL 2605 to (0, -21, 2.2) mm, rotated rx 0 ry 0 rz 180 deg; joints [18.113, -54.782, 108.382, -157.883, 55.667, 77.09]
  MoveL 2606 to (-200, -21, 2.2) mm, rotated rx 0 ry 0 rz 180 deg; joints [20.954, -63.819, 124.325, -156.253, 62.627, 78.565]
  MoveL 2607 to (-200, -21.6, 2.2) mm, rotated rx 0 ry 0 rz 180 deg; joints [20.954, -63.853, 124.319, -156.245, 62.59, 78.546]
  MoveL 2608 to (0, -21.6, 2.2) mm, rotated rx 0 ry 0 rz 180 deg; joints [18.113, -54.81, 108.376, -157.874, 55.635, 77.075]
  MoveL 2609 to (0, -22.2, 2.2) mm, rotated rx 0 ry 0 rz 180 deg; joints [18.113, -54.838, 108.37, -157.866, 55.603, 77.059]
  MoveL 2610 to (-200, -22.2, 2.2) mm, rotated rx 0 ry 0 rz 180 deg; joints [20.954, -63.887, 124.312, -156.236, 62.553, 78.528]
  MoveL 2611 to (-200, -22.8, 2.2) mm, rotated rx 0 ry 0 rz 180 deg; joints [20.954, -63.922, 124.306, -156.227, 62.516, 78.509]
  MoveL 2612 to (0, -22.8, 2.2) mm, rotated rx 0 ry 0 rz 180 deg; joints [18.113, -54.866, 108.364, -157.857, 55.572, 77.043]
  MoveL 2613 to (0, -23.4, 2.2) mm, rotated rx 0 ry 0 rz 180 deg; joints [18.113, -54.895, 108.358, -157.848, 55.54, 77.028]
  MoveL 2614 to (-200, -23.4, 2.2) mm, rotated rx 0 ry 0 rz 180 deg; joints [20.954, -63.956, 124.299, -156.219, 62.478, 78.491]
  MoveL 2615 to (-200, -24, 2.2) mm, rotated rx 0 ry 0 rz 180 deg; joints [20.954, -63.99, 124.292, -156.21, 62.441, 78.472]
  MoveL 2616 to (0, -24, 2.2) mm, rotated rx 0 ry 0 rz 180 deg; joints [18.113, -54.923, 108.352, -157.839, 55.509, 77.012]
  MoveL 2617 to (0, -24.6, 2.2) mm, rotated rx 0 ry 0 rz 180 deg; joints [18.113, -54.951, 108.346, -157.83, 55.477, 76.997]
  MoveL 2618 to (-200, -24.6, 2.2) mm, rotated rx 0 ry 0 rz 180 deg; joints [20.954, -64.024, 124.286, -156.202, 62.404, 78.454]
  MoveL 2619 to (-200, -25.2, 2.2) mm, rotated rx 0 ry 0 rz 180 deg; joints [20.954, -64.058, 124.279, -156.193, 62.367, 78.435]
  MoveL 2620 to (0, -25.2, 2.2) mm, rotated rx 0 ry 0 rz 180 deg; joints [18.113, -54.979, 108.34, -157.821, 55.445, 76.981]
  MoveL 2621 to (0, -25.8, 2.2) mm, rotated rx 0 ry 0 rz 180 deg; joints [18.113, -55.007, 108.334, -157.812, 55.414, 76.965]
  MoveL 2622 to (-200, -25.8, 2.2) mm, rotated rx 0 ry 0 rz 180 deg; joints [20.954, -64.092, 124.273, -156.185, 62.33, 78.417]
  MoveL 2623 to (-200, -26.4, 2.2) mm, rotated rx 0 ry 0 rz 180 deg; joints [20.954, -64.126, 124.266, -156.176, 62.292, 78.398]
  MoveL 2624 to (0, -26.4, 2.2) mm, rotated rx 0 ry 0 rz 180 deg; joints [18.113, -55.035, 108.328, -157.804, 55.382, 76.95]
  MoveL 2625 to (0, -27, 2.2) mm, rotated rx 0 ry 0 rz 180 deg; joints [18.113, -55.063, 108.322, -157.795, 55.35, 76.934]
  MoveL 2626 to (-200, -27, 2.2) mm, rotated rx 0 ry 0 rz 180 deg; joints [20.954, -64.16, 124.259, -156.167, 62.255, 78.379]
  MoveL 2627 to (-200, -27.6, 2.2) mm, rotated rx 0 ry 0 rz 180 deg; joints [20.954, -64.194, 124.252, -156.159, 62.218, 78.361]
  MoveL 2628 to (0, -27.6, 2.2) mm, rotated rx 0 ry 0 rz 180 deg; joints [18.113, -55.091, 108.315, -157.786, 55.319, 76.918]
  MoveL 2629 to (0, -28.2, 2.2) mm, rotated rx 0 ry 0 rz 180 deg; joints [18.113, -55.119, 108.309, -157.777, 55.287, 76.902]
  MoveL 2630 to (-200, -28.2, 2.2) mm, rotated rx 0 ry 0 rz 180 deg; joints [20.954, -64.228, 124.246, -156.15, 62.18, 78.342]
  MoveL 2631 to (-200, -28.8, 2.2) mm, rotated rx 0 ry 0 rz 180 deg; joints [20.954, -64.262, 124.239, -156.141, 62.143, 78.324]
  MoveL 2632 to (0, -28.8, 2.2) mm, rotated rx 0 ry 0 rz 180 deg; joints [18.113, -55.147, 108.303, -157.768, 55.255, 76.887]
  MoveL 2633 to (0, -29.4, 2.2) mm, rotated rx 0 ry 0 rz 180 deg; joints [18.113, -55.175, 108.297, -157.759, 55.224, 76.871]
  MoveL 2634 to (-200, -29.4, 2.2) mm, rotated rx 0 ry 0 rz 180 deg; joints [20.954, -64.296, 124.232, -156.133, 62.106, 78.305]
  MoveL 2635 to (-200, -30, 2.2) mm, rotated rx 0 ry 0 rz 180 deg; joints [20.954, -64.33, 124.225, -156.124, 62.069, 78.286]
  MoveL 2636 to (0, -30, 2.2) mm, rotated rx 0 ry 0 rz 180 deg; joints [18.113, -55.203, 108.29, -157.75, 55.192, 76.855]
  MoveL 2637 to (0, -30.6, 2.21) mm, rotated rx 2.69 ry 0 rz 180 deg; joints [18.022, -56.038, 108.162, -157.6, 54.279, 79.156]
  MoveL 2638 to (-200, -30.6, 2.21) mm, rotated rx 2.69 ry 0 rz 180 deg; joints [20.85, -65.341, 124.083, -155.985, 60.993, 80.495]
  MoveL 2639 to (-200, -31.2, 2.26) mm, rotated rx 5.37 ry 0 rz 180 deg; joints [20.711, -66.341, 123.938, -155.876, 59.918, 82.72]
  MoveL 2640 to (0, -31.2, 2.26) mm, rotated rx 5.37 ry 0 rz 180 deg; joints [17.899, -56.866, 108.033, -157.48, 53.367, 81.475]
  MoveL 2641 to (0, -31.79, 2.33) mm, rotated rx 8.06 ry 0 rz 180 deg; joints [17.746, -57.684, 107.904, -157.392, 52.454, 83.818]
  MoveL 2642 to (-200, -31.79, 2.33) mm, rotated rx 8.06 ry 0 rz 180 deg; joints [20.538, -67.33, 123.792, -155.797, 58.844, 84.966]
  MoveL 2643 to (-200, -32.39, 2.42) mm, rotated rx 10.74 ry 0 rz 180 deg; joints [20.331, -68.304, 123.646, -155.751, 57.774, 87.236]
  MoveL 2644 to (0, -32.39, 2.42) mm, rotated rx 10.74 ry 0 rz 180 deg; joints [17.563, -58.491, 107.774, -157.335, 51.544, 86.185]
  MoveL 2645 to (0, -32.97, 2.55) mm, rotated rx 13.43 ry 0 rz 180 deg; joints [17.35, -59.286, 107.646, -157.313, 50.638, 88.58]
  MoveL 2646 to (-200, -32.97, 2.55) mm, rotated rx 13.43 ry 0 rz 180 deg; joints [20.089, -69.263, 123.498, -155.738, 56.709, 89.533]
  MoveL 2647 to (-200, -33.55, 2.7) mm, rotated rx 16.11 ry 0 rz 180 deg; joints [19.813, -70.203, 123.351, -155.761, 55.65, 91.86]
  MoveL 2648 to (0, -33.55, 2.7) mm, rotated rx 16.11 ry 0 rz 180 deg; joints [17.106, -60.067, 107.518, -157.327, 49.737, 91.005]
  MoveL 2649 to (0, -34.12, 2.88) mm, rotated rx 18.8 ry 0 rz 180 deg; joints [16.833, -60.832, 107.392, -157.379, 48.842, 93.464]
  MoveL 2650 to (-200, -34.12, 2.88) mm, rotated rx 18.8 ry 0 rz 180 deg; joints [19.504, -71.125, 123.205, -155.821, 54.599, 94.221]
  MoveL 2651 to (-200, -34.69, 3.09) mm, rotated rx 21.49 ry 0 rz 180 deg; joints [19.16, -72.027, 123.061, -155.921, 53.557, 96.619]
  MoveL 2652 to (0, -34.69, 3.09) mm, rotated rx 21.49 ry 0 rz 180 deg; joints [16.531, -61.581, 107.268, -157.471, 47.955, 95.96]
  MoveL 2653 to (0, -35.24, 3.32) mm, rotated rx 24.17 ry 0 rz 180 deg; joints [16.201, -62.312, 107.146, -157.604, 47.079, 98.497]
  MoveL 2654 to (-200, -35.24, 3.32) mm, rotated rx 24.17 ry 0 rz 180 deg; joints [18.784, -72.906, 122.919, -156.063, 52.527, 99.059]
  MoveL 2655 to (-200, -35.78, 3.58) mm, rotated rx 26.86 ry 0 rz 180 deg; joints [18.376, -73.761, 122.78, -156.249, 51.51, 101.541]
  MoveL 2656 to (0, -35.78, 3.58) mm, rotated rx 26.86 ry 0 rz 180 deg; joints [15.842, -63.024, 107.028, -157.782, 46.214, 101.075]
  MoveL 2657 to (0, -36.31, 3.86) mm, rotated rx 29.54 ry 0 rz 180 deg; joints [15.455, -63.715, 106.914, -158.007, 45.362, 103.7]
  MoveL 2658 to (-200, -36.31, 3.86) mm, rotated rx 29.54 ry 0 rz 180 deg; joints [17.935, -74.592, 122.644, -156.483, 50.508, 104.073]
  MoveL 2659 to (-200, -36.83, 4.17) mm, rotated rx 32.23 ry 0 rz 180 deg; joints [17.462, -75.396, 122.513, -156.766, 49.523, 106.657]
  MoveL 2660 to (0, -36.83, 4.17) mm, rotated rx 32.23 ry 0 rz 180 deg; joints [15.041, -64.385, 106.805, -158.28, 44.526, 106.375]
  MoveL 2661 to (0, -37.33, 4.5) mm, rotated rx 34.92 ry 0 rz 180 deg; joints [14.6, -65.031, 106.701, -158.605, 43.708, 109.102]
  MoveL 2662 to (-200, -37.33, 4.5) mm, rotated rx 34.92 ry 0 rz 180 deg; joints [16.958, -76.172, 122.387, -157.102, 48.558, 109.296]
  MoveL 2663 to (-200, -37.81, 4.86) mm, rotated rx 37.6 ry 0 rz 180 deg; joints [16.424, -76.919, 122.268, -157.492, 47.614, 111.993]
  MoveL 2664 to (0, -37.81, 4.86) mm, rotated rx 37.6 ry 0 rz 180 deg; joints [14.134, -65.653, 106.603, -158.983, 42.91, 111.883]
  MoveL 2665 to (0, -38.28, 5.24) mm, rotated rx 40.29 ry 0 rz 180 deg; joints [13.642, -66.251, 106.511, -159.416, 42.133, 114.723]
  MoveL 2666 to (-200, -38.28, 5.24) mm, rotated rx 40.29 ry 0 rz 180 deg; joints [15.861, -77.636, 122.155, -157.941, 46.695, 114.753]
  MoveL 2667 to (-200, -38.73, 5.63) mm, rotated rx 42.97 ry 0 rz 180 deg; joints [15.269, -78.322, 122.049, -158.449, 45.803, 117.579]
  MoveL 2668 to (0, -38.73, 5.63) mm, rotated rx 42.97 ry 0 rz 180 deg; joints [13.126, -66.822, 106.426, -159.907, 41.381, 117.624]
  MoveL 2669 to (0, -39.15, 6.05) mm, rotated rx 45.66 ry 0 rz 180 deg; joints [12.587, -67.366, 106.349, -160.458, 40.655, 120.587]
  MoveL 2670 to (-200, -39.15, 6.05) mm, rotated rx 45.66 ry 0 rz 180 deg; joints [14.649, -78.974, 121.952, -159.021, 44.941, 120.473]
  MoveL 2671 to (-200, -39.56, 6.49) mm, rotated rx 48.34 ry 0 rz 180 deg; joints [14.003, -79.593, 121.864, -159.657, 44.112, 123.437]
  MoveL 2672 to (0, -39.56, 6.49) mm, rotated rx 48.34 ry 0 rz 180 deg; joints [12.026, -67.881, 106.281, -161.07, 39.96, 123.614]
  MoveL 2673 to (0, -39.95, 6.95) mm, rotated rx 51.03 ry 0 rz 180 deg; joints [11.444, -68.368, 106.221, -161.744, 39.296, 126.708]
  MoveL 2674 to (-200, -39.95, 6.95) mm, rotated rx 51.03 ry 0 rz 180 deg; joints [13.332, -80.176, 121.786, -160.361, 43.319, 126.475]
  MoveL 2675 to (-200, -40.32, 7.42) mm, rotated rx 53.72 ry 0 rz 180 deg; joints [12.636, -80.724, 121.718, -161.132, 42.565, 129.587]
  MoveL 2676 to (0, -40.32, 7.42) mm, rotated rx 53.72 ry 0 rz 180 deg; joints [10.841, -68.824, 106.171, -162.48, 38.667, 129.869]
  MoveL 2677 to (0, -40.66, 7.92) mm, rotated rx 56.4 ry 0 rz 180 deg; joints [10.219, -69.25, 106.131, -163.28, 38.076, 133.097]
  MoveL 2678 to (-200, -40.66, 7.92) mm, rotated rx 56.4 ry 0 rz 180 deg; joints [11.917, -81.235, 121.661, -161.972, 41.854, 132.775]
  MoveL 2679 to (-200, -40.98, 8.42) mm, rotated rx 59.09 ry 0 rz 180 deg; joints [11.177, -81.708, 121.615, -162.881, 41.19, 136.036]
  MoveL 2680 to (0, -40.98, 8.42) mm, rotated rx 59.09 ry 0 rz 180 deg; joints [9.581, -69.644, 106.101, -164.143, 37.526, 136.391]
  MoveL 2681 to (0, -41.28, 8.95) mm, rotated rx 61.77 ry 0 rz 180 deg; joints [8.926, -70.005, 106.082, -165.067, 37.019, 139.751]
  MoveL 2682 to (-200, -41.28, 8.95) mm, rotated rx 61.77 ry 0 rz 180 deg; joints [10.418, -82.142, 121.582, -163.859, 40.575, 139.374]
  MoveL 2683 to (-200, -41.55, 9.48) mm, rotated rx 64.46 ry 0 rz 180 deg; joints [9.64, -82.536, 121.561, -164.903, 40.013, 142.784]
  MoveL 2684 to (0, -41.55, 9.48) mm, rotated rx 64.46 ry 0 rz 180 deg; joints [8.256, -70.333, 106.075, -166.05, 36.558, 143.174]
  MoveL 2685 to (0, -41.8, 10.03) mm, rotated rx 67.14 ry 0 rz 180 deg; joints [7.573, -70.628, 106.078, -167.089, 36.147, 146.656]
  MoveL 2686 to (-200, -41.8, 10.03) mm, rotated rx 67.14 ry 0 rz 180 deg; joints [8.847, -82.89, 121.554, -166.011, 39.508, 146.263]
  MoveL 2687 to (-200, -42.02, 10.59) mm, rotated rx 69.83 ry 0 rz 180 deg; joints [8.038, -83.203, 121.56, -167.179, 39.062, 149.808]
  MoveL 2688 to (0, -42.02, 10.59) mm, rotated rx 69.83 ry 0 rz 180 deg; joints [6.879, -70.888, 106.094, -168.182, 35.787, 150.195]
  MoveL 2689 to (0, -42.21, 11.15) mm, rotated rx 72.52 ry 0 rz 180 deg; joints [6.174, -71.113, 106.122, -169.322, 35.48, 153.785]
  MoveL 2690 to (-200, -42.21, 11.15) mm, rotated rx 72.52 ry 0 rz 180 deg; joints [7.217, -83.475, 121.58, -168.403, 38.68, 153.413]
  MoveL 2691 to (-200, -42.38, 11.73) mm, rotated rx 75.2 ry 0 rz 180 deg; joints [6.386, -83.703, 121.613, -169.676, 38.364, 157.072]
  MoveL 2692 to (0, -42.38, 11.73) mm, rotated rx 75.2 ry 0 rz 180 deg; joints [5.461, -71.303, 106.162, -170.504, 35.231, 157.42]
  MoveL 2693 to (0, -42.52, 12.31) mm, rotated rx 77.89 ry 0 rz 180 deg; joints [4.742, -71.457, 106.214, -171.72, 35.039, 161.091]
  MoveL 2694 to (-200, -42.52, 12.31) mm, rotated rx 77.89 ry 0 rz 180 deg; joints [5.547, -83.889, 121.661, -170.99, 38.117, 160.775]
  MoveL 2695 to (-200, -42.63, 12.9) mm, rotated rx 80.57 ry 0 rz 180 deg; joints [4.701, -84.031, 121.723, -172.339, 37.941, 164.517]
  MoveL 2696 to (0, -42.63, 12.9) mm, rotated rx 80.57 ry 0 rz 180 deg; joints [4.018, -71.574, 106.278, -172.966, 34.907, 164.794]
  MoveL 2697 to (0, -42.71, 13.5) mm, rotated rx 83.26 ry 0 rz 180 deg; joints [3.292, -71.655, 106.355, -174.231, 34.836, 168.518]
  MoveL 2698 to (-200, -42.71, 13.5) mm, rotated rx 83.26 ry 0 rz 180 deg; joints [3.852, -84.13, 121.799, -173.713, 37.837, 168.285]
  MoveL 2699 to (-200, -42.77, 14.1) mm, rotated rx 85.94 ry 0 rz 180 deg; joints [3, -84.184, 121.89, -175.102, 37.807, 172.071]
  MoveL 2700 to (0, -42.77, 14.1) mm, rotated rx 85.94 ry 0 rz 180 deg; joints [2.563, -71.7, 106.444, -175.508, 34.827, 172.254]
  MoveL 2701 to (0, -42.8, 14.69) mm, rotated rx 88.63 ry 0 rz 180 deg; joints [1.836, -71.707, 106.544, -176.788, 34.88, 175.993]
  MoveL 2702 to (-200, -42.8, 14.69) mm, rotated rx 88.63 ry 0 rz 180 deg; joints [2.15, -84.194, 121.994, -176.496, 37.852, 175.861]
  MoveL 2703 to (-200, -42.8, 15.29) mm, rotated rx 90 ry 0 rz 180 deg; joints [1.702, -84.182, 122.053, -177.229, 37.903, 177.813]
  MoveL 2704 to (0, -42.8, 15.29) mm, rotated rx 90 ry 0 rz 180 deg; joints [1.454, -71.696, 106.601, -177.46, 34.931, 177.918]
  MoveL 2705 to (0, -42.8, 15.89) mm, rotated rx 90 ry 0 rz 180 deg; joints [1.429, -71.697, 106.602, -177.504, 34.93, 177.953]
  MoveL 2706 to (-200, -42.8, 15.89) mm, rotated rx 90 ry 0 rz 180 deg; joints [1.672, -84.183, 122.054, -177.277, 37.902, 177.851]
  MoveL 2707 to (-200, -42.8, 16.49) mm, rotated rx 90 ry 0 rz 180 deg; joints [1.643, -84.185, 122.056, -177.325, 37.901, 177.888]
  MoveL 2708 to (0, -42.8, 16.49) mm, rotated rx 90 ry 0 rz 180 deg; joints [1.404, -71.698, 106.603, -177.548, 34.93, 177.989]
  MoveL 2709 to (0, -42.8, 17.09) mm, rotated rx 90 ry 0 rz 180 deg; joints [1.379, -71.699, 106.605, -177.592, 34.929, 178.025]
  MoveL 2710 to (-200, -42.8, 17.09) mm, rotated rx 90 ry 0 rz 180 deg; joints [1.614, -84.186, 122.057, -177.372, 37.901, 177.926]
  MoveL 2711 to (-200, -42.8, 17.69) mm, rotated rx 90 ry 0 rz 180 deg; joints [1.585, -84.187, 122.058, -177.42, 37.9, 177.964]
  MoveL 2712 to (0, -42.8, 17.69) mm, rotated rx 90 ry 0 rz 180 deg; joints [1.354, -71.7, 106.606, -177.635, 34.929, 178.061]
  MoveL 2713 to (0, -42.8, 18.29) mm, rotated rx 90 ry 0 rz 180 deg; joints [1.329, -71.701, 106.607, -177.679, 34.928, 178.097]
  MoveL 2714 to (-200, -42.8, 18.29) mm, rotated rx 90 ry 0 rz 180 deg; joints [1.555, -84.188, 122.059, -177.468, 37.899, 178.001]
  MoveL 2715 to (-200, -42.8, 18.89) mm, rotated rx 90 ry 0 rz 180 deg; joints [1.526, -84.189, 122.06, -177.515, 37.898, 178.039]
  MoveL 2716 to (0, -42.8, 18.89) mm, rotated rx 90 ry 0 rz 180 deg; joints [1.304, -71.702, 106.608, -177.723, 34.928, 178.133]
  MoveL 2717 to (0, -42.8, 19.49) mm, rotated rx 90 ry 0 rz 180 deg; joints [1.278, -71.703, 106.609, -177.767, 34.927, 178.169]
  MoveL 2718 to (-200, -42.8, 19.49) mm, rotated rx 90 ry 0 rz 180 deg; joints [1.497, -84.19, 122.062, -177.563, 37.897, 178.077]
  MoveL 2719 to (-200, -42.8, 20.09) mm, rotated rx 90 ry 0 rz 180 deg; joints [1.467, -84.191, 122.063, -177.611, 37.896, 178.114]
  MoveL 2720 to (0, -42.8, 20.09) mm, rotated rx 90 ry 0 rz 180 deg; joints [1.253, -71.703, 106.61, -177.81, 34.927, 178.204]
  MoveL 2721 to (0, -42.8, 20.69) mm, rotated rx 90 ry 0 rz 180 deg; joints [1.228, -71.704, 106.611, -177.854, 34.926, 178.24]
  MoveL 2722 to (-200, -42.8, 20.69) mm, rotated rx 90 ry 0 rz 180 deg; joints [1.438, -84.192, 122.064, -177.658, 37.895, 178.152]
  MoveL 2723 to (-200, -42.8, 21.29) mm, rotated rx 90 ry 0 rz 180 deg; joints [1.409, -84.193, 122.065, -177.706, 37.894, 178.189]
  MoveL 2724 to (0, -42.8, 21.29) mm, rotated rx 90 ry 0 rz 180 deg; joints [1.203, -71.705, 106.613, -177.898, 34.926, 178.276]
  MoveL 2725 to (0, -42.8, 21.89) mm, rotated rx 90 ry 0 rz 180 deg; joints [1.178, -71.706, 106.614, -177.942, 34.925, 178.312]
  MoveL 2726 to (-200, -42.8, 21.89) mm, rotated rx 90 ry 0 rz 180 deg; joints [1.379, -84.194, 122.066, -177.754, 37.894, 178.227]
  MoveL 2727 to (-200, -42.8, 22.49) mm, rotated rx 90 ry 0 rz 180 deg; joints [1.35, -84.195, 122.067, -177.802, 37.893, 178.265]
  MoveL 2728 to (0, -42.8, 22.49) mm, rotated rx 90 ry 0 rz 180 deg; joints [1.153, -71.707, 106.615, -177.985, 34.925, 178.348]
  MoveL 2729 to (0, -42.8, 23.09) mm, rotated rx 90 ry 0 rz 180 deg; joints [1.128, -71.707, 106.616, -178.029, 34.924, 178.384]
  MoveL 2730 to (-200, -42.8, 23.09) mm, rotated rx 90 ry 0 rz 180 deg; joints [1.321, -84.196, 122.068, -177.849, 37.892, 178.302]
  MoveL 2731 to (-200, -42.8, 23.69) mm, rotated rx 90 ry 0 rz 180 deg; joints [1.291, -84.196, 122.069, -177.897, 37.891, 178.34]
  MoveL 2732 to (0, -42.8, 23.69) mm, rotated rx 90 ry 0 rz 180 deg; joints [1.103, -71.708, 106.617, -178.073, 34.924, 178.42]
  MoveL 2733 to (0, -42.8, 24.29) mm, rotated rx 90 ry 0 rz 180 deg; joints [1.078, -71.709, 106.617, -178.117, 34.923, 178.456]
  MoveL 2734 to (-200, -42.8, 24.29) mm, rotated rx 90 ry 0 rz 180 deg; joints [1.262, -84.197, 122.07, -177.945, 37.891, 178.378]
  MoveL 2735 to (-200, -42.8, 24.89) mm, rotated rx 90 ry 0 rz 180 deg; joints [1.233, -84.198, 122.071, -177.993, 37.89, 178.415]
  MoveL 2736 to (0, -42.8, 24.89) mm, rotated rx 90 ry 0 rz 180 deg; joints [1.053, -71.709, 106.618, -178.16, 34.923, 178.491]
  MoveL 2737 to (0, -42.8, 25.49) mm, rotated rx 90 ry 0 rz 180 deg; joints [1.028, -71.71, 106.619, -178.204, 34.922, 178.527]
  MoveL 2738 to (-200, -42.8, 25.49) mm, rotated rx 90 ry 0 rz 180 deg; joints [1.203, -84.199, 122.072, -178.04, 37.889, 178.453]
  MoveL 2739 to (-200, -42.8, 26.09) mm, rotated rx 90 ry 0 rz 180 deg; joints [1.174, -84.2, 122.073, -178.088, 37.888, 178.491]
  MoveL 2740 to (0, -42.8, 26.09) mm, rotated rx 90 ry 0 rz 180 deg; joints [1.003, -71.711, 106.62, -178.248, 34.922, 178.563]
  MoveL 2741 to (0, -42.8, 26.69) mm, rotated rx 90 ry 0 rz 180 deg; joints [0.978, -71.711, 106.621, -178.292, 34.922, 178.599]
  MoveL 2742 to (-200, -42.8, 26.69) mm, rotated rx 90 ry 0 rz 180 deg; joints [1.145, -84.2, 122.074, -178.136, 37.888, 178.528]
  MoveL 2743 to (-200, -42.8, 27.29) mm, rotated rx 90 ry 0 rz 180 deg; joints [1.115, -84.201, 122.074, -178.183, 37.887, 178.566]
  MoveL 2744 to (0, -42.8, 27.29) mm, rotated rx 90 ry 0 rz 180 deg; joints [0.953, -71.712, 106.622, -178.335, 34.921, 178.635]
  MoveL 2745 to (0, -42.8, 27.89) mm, rotated rx 90 ry 0 rz 180 deg; joints [0.928, -71.713, 106.623, -178.379, 34.921, 178.671]
  MoveL 2746 to (-200, -42.8, 27.89) mm, rotated rx 90 ry 0 rz 180 deg; joints [1.086, -84.202, 122.075, -178.231, 37.886, 178.604]
  MoveL 2747 to (-200, -42.8, 28.49) mm, rotated rx 90 ry 0 rz 180 deg; joints [1.057, -84.203, 122.076, -178.279, 37.886, 178.641]
  MoveL 2748 to (0, -42.8, 28.49) mm, rotated rx 90 ry 0 rz 180 deg; joints [0.903, -71.713, 106.624, -178.423, 34.921, 178.707]
  MoveL 2749 to (0, -42.8, 29.09) mm, rotated rx 90 ry 0 rz 180 deg; joints [0.878, -71.714, 106.624, -178.467, 34.92, 178.743]
  MoveL 2750 to (-200, -42.8, 29.09) mm, rotated rx 90 ry 0 rz 180 deg; joints [1.027, -84.203, 122.077, -178.327, 37.885, 178.679]
  MoveL 2751 to (-200, -42.8, 29.69) mm, rotated rx 90 ry 0 rz 180 deg; joints [0.998, -84.204, 122.078, -178.374, 37.885, 178.717]
  MoveL 2752 to (0, -42.8, 29.69) mm, rotated rx 90 ry 0 rz 180 deg; joints [0.853, -71.714, 106.625, -178.51, 34.92, 178.778]
  MoveL 2753 to (0, -42.8, 30.29) mm, rotated rx 90 ry 0 rz 180 deg; joints [0.828, -71.715, 106.626, -178.554, 34.92, 178.814]
  MoveL 2754 to (-200, -42.8, 30.29) mm, rotated rx 90 ry 0 rz 180 deg; joints [0.969, -84.205, 122.078, -178.422, 37.884, 178.755]
  MoveL 2755 to (-200, -42.8, 30.89) mm, rotated rx 90 ry 0 rz 180 deg; joints [0.94, -84.205, 122.079, -178.47, 37.884, 178.792]
  MoveL 2756 to (0, -42.8, 30.89) mm, rotated rx 90 ry 0 rz 180 deg; joints [0.803, -71.715, 106.627, -178.598, 34.919, 178.85]
  MoveL 2757 to (0, -42.8, 31.49) mm, rotated rx 90 ry 0 rz 180 deg; joints [0.778, -71.716, 106.627, -178.642, 34.919, 178.886]
  MoveL 2758 to (-200, -42.8, 31.49) mm, rotated rx 90 ry 0 rz 180 deg; joints [0.91, -84.206, 122.08, -178.518, 37.883, 178.83]
  MoveL 2759 to (-200, -42.8, 32.09) mm, rotated rx 90 ry 0 rz 180 deg; joints [0.881, -84.207, 122.08, -178.565, 37.882, 178.868]
  MoveL 2760 to (0, -42.8, 32.09) mm, rotated rx 90 ry 0 rz 180 deg; joints [0.752, -71.716, 106.628, -178.685, 34.919, 178.922]
  MoveL 2761 to (0, -42.8, 32.69) mm, rotated rx 90 ry 0 rz 180 deg; joints [0.727, -71.717, 106.629, -178.729, 34.918, 178.958]
  MoveL 2762 to (-200, -42.8, 32.69) mm, rotated rx 90 ry 0 rz 180 deg; joints [0.852, -84.207, 122.081, -178.613, 37.882, 178.905]
  MoveL 2763 to (-200, -42.8, 33.29) mm, rotated rx 90 ry 0 rz 180 deg; joints [0.822, -84.208, 122.082, -178.661, 37.881, 178.943]
  MoveL 2764 to (0, -42.8, 33.29) mm, rotated rx 90 ry 0 rz 180 deg; joints [0.702, -71.717, 106.629, -178.773, 34.918, 178.994]
  MoveL 2765 to (0, -42.8, 33.89) mm, rotated rx 90 ry 0 rz 180 deg; joints [0.677, -71.718, 106.63, -178.817, 34.918, 179.03]
  MoveL 2766 to (-200, -42.8, 33.89) mm, rotated rx 90 ry 0 rz 180 deg; joints [0.793, -84.208, 122.082, -178.709, 37.881, 178.981]
  MoveL 2767 to (-200, -42.8, 34.49) mm, rotated rx 90 ry 0 rz 180 deg; joints [0.764, -84.209, 122.083, -178.756, 37.881, 179.018]
  MoveL 2768 to (0, -42.8, 34.49) mm, rotated rx 90 ry 0 rz 180 deg; joints [0.652, -71.718, 106.63, -178.86, 34.917, 179.066]
  MoveL 2769 to (0, -42.8, 35.09) mm, rotated rx 90 ry 0 rz 180 deg; joints [0.627, -71.719, 106.631, -178.904, 34.917, 179.101]
  MoveL 2770 to (-200, -42.8, 35.09) mm, rotated rx 90 ry 0 rz 180 deg; joints [0.734, -84.209, 122.083, -178.804, 37.88, 179.056]
  MoveL 2771 to (-200, -42.8, 35.69) mm, rotated rx 90 ry 0 rz 180 deg; joints [0.705, -84.21, 122.084, -178.852, 37.88, 179.094]
  MoveL 2772 to (0, -42.8, 35.69) mm, rotated rx 90 ry 0 rz 180 deg; joints [0.602, -71.719, 106.631, -178.948, 34.917, 179.137]
  MoveL 2773 to (0, -42.8, 36.29) mm, rotated rx 90 ry 0 rz 180 deg; joints [0.577, -71.719, 106.632, -178.992, 34.917, 179.173]
  MoveL 2774 to (-200, -42.8, 36.29) mm, rotated rx 90 ry 0 rz 180 deg; joints [0.676, -84.21, 122.084, -178.9, 37.879, 179.131]
  MoveL 2775 to (-200, -42.8, 36.89) mm, rotated rx 90 ry 0 rz 180 deg; joints [0.646, -84.211, 122.085, -178.947, 37.879, 179.169]
  MoveL 2776 to (0, -42.8, 36.89) mm, rotated rx 90 ry 0 rz 180 deg; joints [0.552, -71.72, 106.632, -179.036, 34.916, 179.209]
  MoveL 2777 to (0, -42.8, 37.49) mm, rotated rx 90 ry 0 rz 180 deg; joints [0.527, -71.72, 106.633, -179.079, 34.916, 179.245]
  MoveL 2778 to (-200, -42.8, 37.49) mm, rotated rx 90 ry 0 rz 180 deg; joints [0.617, -84.211, 122.085, -178.995, 37.879, 179.207]
  MoveL 2779 to (-200, -42.8, 38.09) mm, rotated rx 90 ry 0 rz 180 deg; joints [0.588, -84.212, 122.086, -179.043, 37.878, 179.245]
  MoveL 2780 to (0, -42.8, 38.09) mm, rotated rx 90 ry 0 rz 180 deg; joints [0.502, -71.72, 106.633, -179.123, 34.916, 179.281]
  MoveL 2781 to (0, -42.8, 38.69) mm, rotated rx 90 ry 0 rz 180 deg; joints [0.477, -71.721, 106.634, -179.167, 34.916, 179.317]
  MoveL 2782 to (-200, -42.8, 38.69) mm, rotated rx 90 ry 0 rz 180 deg; joints [0.558, -84.212, 122.086, -179.091, 37.878, 179.282]
  MoveL 2783 to (-200, -42.8, 39.29) mm, rotated rx 90 ry 0 rz 180 deg; joints [0.529, -84.212, 122.087, -179.139, 37.878, 179.32]
  MoveL 2784 to (0, -42.8, 39.29) mm, rotated rx 90 ry 0 rz 180 deg; joints [0.452, -71.721, 106.634, -179.211, 34.916, 179.353]
  MoveL 2785 to (0, -42.8, 39.89) mm, rotated rx 90 ry 0 rz 180 deg; joints [0.427, -71.721, 106.635, -179.254, 34.915, 179.389]
  MoveL 2786 to (-200, -42.8, 39.89) mm, rotated rx 90 ry 0 rz 180 deg; joints [0.5, -84.213, 122.087, -179.186, 37.877, 179.358]
  MoveL 2787 to (-200, -42.8, 40.49) mm, rotated rx 90 ry 0 rz 180 deg; joints [0.47, -84.213, 122.088, -179.234, 37.877, 179.395]
  MoveL 2788 to (0, -42.8, 40.49) mm, rotated rx 90 ry 0 rz 180 deg; joints [0.402, -71.722, 106.635, -179.298, 34.915, 179.424]
  MoveL 2789 to (0, -42.8, 41.09) mm, rotated rx 90 ry 0 rz 180 deg; joints [0.377, -71.722, 106.635, -179.342, 34.915, 179.46]
  MoveL 2790 to (-200, -42.8, 41.09) mm, rotated rx 90 ry 0 rz 180 deg; joints [0.441, -84.213, 122.088, -179.282, 37.877, 179.433]
  MoveL 2791 to (-200, -42.8, 41.69) mm, rotated rx 90 ry 0 rz 180 deg; joints [0.412, -84.214, 122.088, -179.33, 37.876, 179.471]
  MoveL 2792 to (0, -42.8, 41.69) mm, rotated rx 90 ry 0 rz 180 deg; joints [0.352, -71.722, 106.636, -179.386, 34.915, 179.496]
  MoveL 2793 to (0, -42.8, 42.29) mm, rotated rx 90 ry 0 rz 180 deg; joints [0.327, -71.722, 106.636, -179.429, 34.915, 179.532]
  MoveL 2794 to (-200, -42.8, 42.29) mm, rotated rx 90 ry 0 rz 180 deg; joints [0.382, -84.214, 122.088, -179.377, 37.876, 179.509]
  MoveL 2795 to (-200, -42.8, 42.89) mm, rotated rx 90 ry 0 rz 180 deg; joints [0.353, -84.214, 122.089, -179.425, 37.876, 179.546]
  MoveL 2796 to (0, -42.8, 42.89) mm, rotated rx 90 ry 0 rz 180 deg; joints [0.301, -71.722, 106.636, -179.473, 34.915, 179.568]
  MoveL 2797 to (0, -42.8, 43.49) mm, rotated rx 90 ry 0 rz 180 deg; joints [0.276, -71.723, 106.636, -179.517, 34.915, 179.604]
  MoveL 2798 to (-200, -42.8, 43.49) mm, rotated rx 90 ry 0 rz 180 deg; joints [0.324, -84.214, 122.089, -179.473, 37.876, 179.584]
  MoveL 2799 to (-200, -42.8, 44.09) mm, rotated rx 90 ry 0 rz 180 deg; joints [0.294, -84.215, 122.089, -179.521, 37.876, 179.622]
  MoveL 2800 to (0, -42.8, 44.09) mm, rotated rx 90 ry 0 rz 180 deg; joints [0.251, -71.723, 106.637, -179.561, 34.915, 179.64]
  MoveL 2801 to (0, -42.8, 44.69) mm, rotated rx 90 ry 0 rz 180 deg; joints [0.226, -71.723, 106.637, -179.605, 34.914, 179.676]
  MoveL 2802 to (-200, -42.8, 44.69) mm, rotated rx 90 ry 0 rz 180 deg; joints [0.265, -84.215, 122.089, -179.568, 37.875, 179.659]
  MoveL 2803 to (-200, -42.8, 45.29) mm, rotated rx 91.31 ry 0 rz 180 deg; joints [-0.165, -84.178, 122.133, 179.732, 37.956, -178.473]
  MoveL 2804 to (0, -42.8, 45.29) mm, rotated rx 91.31 ry 0 rz 180 deg; joints [-0.141, -71.692, 106.678, 179.754, 34.986, -178.483]
  MoveL 2805 to (0, -42.77, 45.89) mm, rotated rx 94 ry 0 rz 180 deg; joints [-0.861, -71.602, 106.77, 178.505, 35.177, -174.777]
  MoveL 2806 to (-200, -42.77, 45.89) mm, rotated rx 94 ry 0 rz 180 deg; joints [-1.008, -84.07, 122.233, 178.368, 38.174, -174.716]
  MoveL 2807 to (-200, -42.71, 46.49) mm, rotated rx 96.69 ry 0 rz 180 deg; joints [-1.844, -83.917, 122.346, 177.035, 38.466, -170.991]
  MoveL 2808 to (0, -42.71, 46.49) mm, rotated rx 96.69 ry 0 rz 180 deg; joints [-1.575, -71.474, 106.873, 177.282, 35.43, -171.098]
  MoveL 2809 to (0, -42.63, 47.08) mm, rotated rx 99.37 ry 0 rz 180 deg; joints [-2.281, -71.31, 106.987, 176.094, 35.741, -167.456]
  MoveL 2810 to (-200, -42.63, 47.08) mm, rotated rx 99.37 ry 0 rz 180 deg; joints [-2.669, -83.72, 122.471, 175.74, 38.828, -167.307]
  MoveL 2811 to (-200, -42.52, 47.67) mm, rotated rx 102.06 ry 0 rz 180 deg; joints [-3.483, -83.479, 122.609, 174.492, 39.259, -163.672]
  MoveL 2812 to (0, -42.52, 47.67) mm, rotated rx 102.06 ry 0 rz 180 deg; joints [-2.976, -71.109, 107.112, 174.946, 36.109, -163.855]
  MoveL 2813 to (0, -42.38, 48.26) mm, rotated rx 104.74 ry 0 rz 180 deg; joints [-3.66, -70.871, 107.246, 173.845, 36.533, -160.303]
  MoveL 2814 to (-200, -42.38, 48.26) mm, rotated rx 104.74 ry 0 rz 180 deg; joints [-4.282, -83.194, 122.758, 173.296, 39.757, -160.092]
  MoveL 2815 to (-200, -42.21, 48.83) mm, rotated rx 107.43 ry 0 rz 180 deg; joints [-5.065, -82.865, 122.918, 172.158, 40.318, -156.575]
  MoveL 2816 to (0, -42.21, 48.83) mm, rotated rx 107.43 ry 0 rz 180 deg; joints [-4.33, -70.598, 107.389, 172.795, 37.009, -156.806]
  MoveL 2817 to (0, -42.02, 49.4) mm, rotated rx 110.11 ry 0 rz 180 deg; joints [-4.984, -70.288, 107.541, 171.801, 37.536, -153.367]
  MoveL 2818 to (-200, -42.02, 49.4) mm, rotated rx 110.11 ry 0 rz 180 deg; joints [-5.83, -82.493, 123.088, 171.083, 40.939, -153.125]
  MoveL 2819 to (-200, -41.8, 49.96) mm, rotated rx 112.8 ry 0 rz 180 deg; joints [-6.575, -82.079, 123.267, 170.073, 41.617, -149.745]
  MoveL 2820 to (0, -41.8, 49.96) mm, rotated rx 112.8 ry 0 rz 180 deg; joints [-5.623, -69.944, 107.7, 170.865, 38.111, -149.989]
  MoveL 2821 to (0, -41.55, 50.51) mm, rotated rx 115.49 ry 0 rz 180 deg; joints [-6.243, -69.565, 107.867, 169.99, 38.73, -146.673]
  MoveL 2822 to (-200, -41.55, 50.51) mm, rotated rx 115.49 ry 0 rz 180 deg; joints [-7.298, -81.622, 123.455, 169.13, 42.349, -146.436]
  MoveL 2823 to (-200, -41.28, 51.04) mm, rotated rx 118.17 ry 0 rz 180 deg; joints [-7.998, -81.124, 123.651, 168.257, 43.131, -143.201]
  MoveL 2824 to (0, -41.28, 51.04) mm, rotated rx 118.17 ry 0 rz 180 deg; joints [-6.844, -69.152, 108.04, 169.176, 39.392, -143.422]
  MoveL 2825 to (0, -40.99, 51.56) mm, rotated rx 120.86 ry 0 rz 180 deg; joints [-7.425, -68.705, 108.219, 168.425, 40.093, -140.237]
  MoveL 2826 to (-200, -40.99, 51.56) mm, rotated rx 120.86 ry 0 rz 180 deg; joints [-8.674, -80.585, 123.853, 167.452, 43.96, -140.04]
